    ELSIF ((x0 = FALSE) AND  (x1 = FALSE) AND  (x2 = TRUE) AND  (x3 = TRUE) AND  ( TRUE ) AND  ( TRUE )) OR ((x0 = FALSE) AND  (x1 = TRUE) AND  (x2 = FALSE) AND  (x3 = TRUE) AND  ( TRUE ) AND  ( TRUE )) OR ((x0 = FALSE) AND  (x1 = TRUE) AND  (x2 = TRUE) AND  ( TRUE ) AND  ( TRUE ) AND  ( TRUE )) OR ((x0 = TRUE) AND  ( TRUE ) AND  (x2 = FALSE) AND  (x3 = TRUE) AND  ( TRUE ) AND  ( TRUE )) OR ((x0 = TRUE) AND  ( TRUE ) AND  (x2 = TRUE) AND  ( TRUE ) AND  ( TRUE ) AND  ( TRUE )) THEN 
        cstate98 := 617; y0 := FALSE; y1 := FALSE; y2 := FALSE;  
    ELSIF ((x0 = FALSE) AND  (x1 = TRUE) AND  (x2 = FALSE) AND  (x3 = FALSE) AND  ( TRUE ) AND  (x5 = FALSE)) OR ((x0 = TRUE) AND  ( TRUE ) AND  (x2 = FALSE) AND  (x3 = FALSE) AND  ( TRUE ) AND  (x5 = FALSE)) THEN 
        cstate98 := 3204; y0 := TRUE; y1 := FALSE; y2 := FALSE;  
    ELSIF ((x0 = FALSE) AND  (x1 = TRUE) AND  (x2 = FALSE) AND  (x3 = FALSE) AND  ( TRUE ) AND  (x5 = TRUE)) OR ((x0 = TRUE) AND  ( TRUE ) AND  (x2 = FALSE) AND  (x3 = FALSE) AND  ( TRUE ) AND  (x5 = TRUE)) THEN 
        cstate98 := 1190; y0 := FALSE; y1 := FALSE; y2 := FALSE;  
    END_IF;
2212:
    IF ((x0 = FALSE) AND  (x1 = FALSE) AND  (x2 = FALSE) AND  (x3 = FALSE) AND  ( TRUE ) AND  (x5 = FALSE)) OR ((x0 = FALSE) AND  (x1 = FALSE) AND  (x2 = FALSE) AND  (x3 = TRUE) AND  (x4 = FALSE) AND  (x5 = FALSE)) THEN 
        cstate98 := 2212; y0 := FALSE; y1 := FALSE; y2 := FALSE;  
    ELSIF ((x0 = FALSE) AND  (x1 = FALSE) AND  (x2 = FALSE) AND  (x3 = FALSE) AND  ( TRUE ) AND  (x5 = TRUE)) OR ((x0 = FALSE) AND  (x1 = FALSE) AND  (x2 = FALSE) AND  (x3 = TRUE) AND  (x4 = FALSE) AND  (x5 = TRUE)) THEN 
        cstate98 := 2215; y0 := FALSE; y1 := FALSE; y2 := FALSE;  
    ELSIF ((x0 = FALSE) AND  (x1 = FALSE) AND  (x2 = FALSE) AND  (x3 = TRUE) AND  (x4 = TRUE) AND  (x5 = FALSE)) THEN 
        cstate98 := 236; y0 := FALSE; y1 := FALSE; y2 := TRUE;  
    ELSIF ((x0 = FALSE) AND  (x1 = FALSE) AND  (x2 = FALSE) AND  (x3 = TRUE) AND  (x4 = TRUE) AND  (x5 = TRUE)) THEN 
        cstate98 := 2190; y0 := FALSE; y1 := FALSE; y2 := FALSE;  
    ELSIF ((x0 = FALSE) AND  (x1 = FALSE) AND  (x2 = TRUE) AND  (x3 = FALSE) AND  ( TRUE ) AND  (x5 = FALSE)) THEN 
        cstate98 := 2704; y0 := FALSE; y1 := TRUE; y2 := FALSE;  
    ELSIF ((x0 = FALSE) AND  (x1 = FALSE) AND  (x2 = TRUE) AND  (x3 = FALSE) AND  ( TRUE ) AND  (x5 = TRUE)) THEN 
        cstate98 := 1714; y0 := FALSE; y1 := FALSE; y2 := FALSE;  
    ELSIF ((x0 = FALSE) AND  (x1 = FALSE) AND  (x2 = TRUE) AND  (x3 = TRUE) AND  ( TRUE ) AND  ( TRUE )) OR ((x0 = FALSE) AND  (x1 = TRUE) AND  (x2 = FALSE) AND  (x3 = TRUE) AND  ( TRUE ) AND  ( TRUE )) OR ((x0 = FALSE) AND  (x1 = TRUE) AND  (x2 = TRUE) AND  ( TRUE ) AND  ( TRUE ) AND  ( TRUE )) OR ((x0 = TRUE) AND  ( TRUE ) AND  (x2 = FALSE) AND  (x3 = TRUE) AND  ( TRUE ) AND  ( TRUE )) OR ((x0 = TRUE) AND  ( TRUE ) AND  (x2 = TRUE) AND  ( TRUE ) AND  ( TRUE ) AND  ( TRUE )) THEN 
        cstate98 := 617; y0 := FALSE; y1 := FALSE; y2 := FALSE;  
    ELSIF ((x0 = FALSE) AND  (x1 = TRUE) AND  (x2 = FALSE) AND  (x3 = FALSE) AND  ( TRUE ) AND  (x5 = FALSE)) OR ((x0 = TRUE) AND  ( TRUE ) AND  (x2 = FALSE) AND  (x3 = FALSE) AND  ( TRUE ) AND  (x5 = FALSE)) THEN 
        cstate98 := 3204; y0 := TRUE; y1 := FALSE; y2 := FALSE;  
    ELSIF ((x0 = FALSE) AND  (x1 = TRUE) AND  (x2 = FALSE) AND  (x3 = FALSE) AND  ( TRUE ) AND  (x5 = TRUE)) OR ((x0 = TRUE) AND  ( TRUE ) AND  (x2 = FALSE) AND  (x3 = FALSE) AND  ( TRUE ) AND  (x5 = TRUE)) THEN 
        cstate98 := 1190; y0 := FALSE; y1 := FALSE; y2 := FALSE;  
    END_IF;
236:
    IF ((x0 = FALSE) AND  (x1 = FALSE) AND  (x2 = FALSE) AND  (x3 = FALSE) AND  ( TRUE ) AND  (x5 = FALSE)) OR ((x0 = FALSE) AND  (x1 = FALSE) AND  (x2 = FALSE) AND  (x3 = TRUE) AND  (x4 = FALSE) AND  (x5 = FALSE)) OR ((x0 = FALSE) AND  (x1 = TRUE) AND  (x2 = FALSE) AND  (x3 = FALSE) AND  ( TRUE ) AND  (x5 = FALSE)) OR ((x0 = TRUE) AND  ( TRUE ) AND  (x2 = FALSE) AND  (x3 = FALSE) AND  ( TRUE ) AND  (x5 = FALSE)) THEN 
        cstate98 := 300; y0 := FALSE; y1 := FALSE; y2 := TRUE;  
    ELSIF ((x0 = FALSE) AND  (x1 = FALSE) AND  (x2 = FALSE) AND  (x3 = FALSE) AND  ( TRUE ) AND  (x5 = TRUE)) OR ((x0 = FALSE) AND  (x1 = FALSE) AND  (x2 = FALSE) AND  (x3 = TRUE) AND  (x4 = FALSE) AND  (x5 = TRUE)) THEN 
        cstate98 := 2223; y0 := FALSE; y1 := FALSE; y2 := FALSE;  
    ELSIF ((x0 = FALSE) AND  (x1 = FALSE) AND  (x2 = FALSE) AND  (x3 = TRUE) AND  (x4 = TRUE) AND  (x5 = FALSE)) THEN 
        cstate98 := 236; y0 := FALSE; y1 := FALSE; y2 := TRUE;  
    ELSIF ((x0 = FALSE) AND  (x1 = FALSE) AND  (x2 = FALSE) AND  (x3 = TRUE) AND  (x4 = TRUE) AND  (x5 = TRUE)) THEN 
        cstate98 := 2190; y0 := FALSE; y1 := FALSE; y2 := FALSE;  
    ELSIF ((x0 = FALSE) AND  (x1 = FALSE) AND  (x2 = TRUE) AND  (x3 = FALSE) AND  ( TRUE ) AND  (x5 = FALSE)) THEN 
        cstate98 := 296; y0 := FALSE; y1 := FALSE; y2 := TRUE;  
    ELSIF ((x0 = FALSE) AND  (x1 = FALSE) AND  (x2 = TRUE) AND  (x3 = FALSE) AND  ( TRUE ) AND  (x5 = TRUE)) THEN 
        cstate98 := 1706; y0 := FALSE; y1 := FALSE; y2 := FALSE;  
    ELSIF ((x0 = FALSE) AND  (x1 = FALSE) AND  (x2 = TRUE) AND  (x3 = TRUE) AND  ( TRUE ) AND  ( TRUE )) OR ((x0 = FALSE) AND  (x1 = TRUE) AND  (x2 = FALSE) AND  (x3 = TRUE) AND  ( TRUE ) AND  ( TRUE )) OR ((x0 = FALSE) AND  (x1 = TRUE) AND  (x2 = TRUE) AND  ( TRUE ) AND  ( TRUE ) AND  ( TRUE )) OR ((x0 = TRUE) AND  ( TRUE ) AND  (x2 = FALSE) AND  (x3 = TRUE) AND  ( TRUE ) AND  ( TRUE )) OR ((x0 = TRUE) AND  ( TRUE ) AND  (x2 = TRUE) AND  ( TRUE ) AND  ( TRUE ) AND  ( TRUE )) THEN 
        cstate98 := 617; y0 := FALSE; y1 := FALSE; y2 := FALSE;  
    ELSIF ((x0 = FALSE) AND  (x1 = TRUE) AND  (x2 = FALSE) AND  (x3 = FALSE) AND  ( TRUE ) AND  (x5 = TRUE)) OR ((x0 = TRUE) AND  ( TRUE ) AND  (x2 = FALSE) AND  (x3 = FALSE) AND  ( TRUE ) AND  (x5 = TRUE)) THEN 
        cstate98 := 1198; y0 := FALSE; y1 := FALSE; y2 := FALSE;  
    END_IF;
2214:
    IF ((x0 = FALSE) AND  (x1 = FALSE) AND  (x2 = FALSE) AND  (x3 = FALSE) AND  ( TRUE ) AND  (x5 = FALSE)) OR ((x0 = FALSE) AND  (x1 = FALSE) AND  (x2 = FALSE) AND  (x3 = TRUE) AND  (x4 = FALSE) AND  (x5 = FALSE)) THEN 
        cstate98 := 2214; y0 := FALSE; y1 := FALSE; y2 := FALSE;  
    ELSIF ((x0 = FALSE) AND  (x1 = FALSE) AND  (x2 = FALSE) AND  (x3 = FALSE) AND  ( TRUE ) AND  (x5 = TRUE)) OR ((x0 = FALSE) AND  (x1 = FALSE) AND  (x2 = FALSE) AND  (x3 = TRUE) AND  (x4 = FALSE) AND  (x5 = TRUE)) THEN 
        cstate98 := 2215; y0 := FALSE; y1 := FALSE; y2 := FALSE;  
    ELSIF ((x0 = FALSE) AND  (x1 = FALSE) AND  (x2 = FALSE) AND  (x3 = TRUE) AND  (x4 = TRUE) AND  (x5 = FALSE)) THEN 
        cstate98 := 238; y0 := FALSE; y1 := FALSE; y2 := TRUE;  
    ELSIF ((x0 = FALSE) AND  (x1 = FALSE) AND  (x2 = FALSE) AND  (x3 = TRUE) AND  (x4 = TRUE) AND  (x5 = TRUE)) THEN 
        cstate98 := 2190; y0 := FALSE; y1 := FALSE; y2 := FALSE;  
    ELSIF ((x0 = FALSE) AND  (x1 = FALSE) AND  (x2 = TRUE) AND  (x3 = FALSE) AND  ( TRUE ) AND  (x5 = FALSE)) THEN 
        cstate98 := 2706; y0 := FALSE; y1 := TRUE; y2 := FALSE;  
    ELSIF ((x0 = FALSE) AND  (x1 = FALSE) AND  (x2 = TRUE) AND  (x3 = FALSE) AND  ( TRUE ) AND  (x5 = TRUE)) THEN 
        cstate98 := 1714; y0 := FALSE; y1 := FALSE; y2 := FALSE;  
    ELSIF ((x0 = FALSE) AND  (x1 = FALSE) AND  (x2 = TRUE) AND  (x3 = TRUE) AND  ( TRUE ) AND  ( TRUE )) OR ((x0 = FALSE) AND  (x1 = TRUE) AND  (x2 = FALSE) AND  (x3 = TRUE) AND  ( TRUE ) AND  ( TRUE )) OR ((x0 = FALSE) AND  (x1 = TRUE) AND  (x2 = TRUE) AND  ( TRUE ) AND  ( TRUE ) AND  ( TRUE )) OR ((x0 = TRUE) AND  ( TRUE ) AND  (x2 = FALSE) AND  (x3 = TRUE) AND  ( TRUE ) AND  ( TRUE )) OR ((x0 = TRUE) AND  ( TRUE ) AND  (x2 = TRUE) AND  ( TRUE ) AND  ( TRUE ) AND  ( TRUE )) THEN 
        cstate98 := 617; y0 := FALSE; y1 := FALSE; y2 := FALSE;  
    ELSIF ((x0 = FALSE) AND  (x1 = TRUE) AND  (x2 = FALSE) AND  (x3 = FALSE) AND  ( TRUE ) AND  (x5 = FALSE)) OR ((x0 = TRUE) AND  ( TRUE ) AND  (x2 = FALSE) AND  (x3 = FALSE) AND  ( TRUE ) AND  (x5 = FALSE)) THEN 
        cstate98 := 3206; y0 := TRUE; y1 := FALSE; y2 := FALSE;  
    ELSIF ((x0 = FALSE) AND  (x1 = TRUE) AND  (x2 = FALSE) AND  (x3 = FALSE) AND  ( TRUE ) AND  (x5 = TRUE)) OR ((x0 = TRUE) AND  ( TRUE ) AND  (x2 = FALSE) AND  (x3 = FALSE) AND  ( TRUE ) AND  (x5 = TRUE)) THEN 
        cstate98 := 1190; y0 := FALSE; y1 := FALSE; y2 := FALSE;  
    END_IF;
238:
    IF ((x0 = FALSE) AND  (x1 = FALSE) AND  (x2 = FALSE) AND  (x3 = FALSE) AND  ( TRUE ) AND  (x5 = FALSE)) OR ((x0 = FALSE) AND  (x1 = FALSE) AND  (x2 = FALSE) AND  (x3 = TRUE) AND  (x4 = FALSE) AND  (x5 = FALSE)) OR ((x0 = FALSE) AND  (x1 = TRUE) AND  (x2 = FALSE) AND  (x3 = FALSE) AND  ( TRUE ) AND  (x5 = FALSE)) OR ((x0 = TRUE) AND  ( TRUE ) AND  (x2 = FALSE) AND  (x3 = FALSE) AND  ( TRUE ) AND  (x5 = FALSE)) THEN 
        cstate98 := 302; y0 := FALSE; y1 := FALSE; y2 := TRUE;  
    ELSIF ((x0 = FALSE) AND  (x1 = FALSE) AND  (x2 = FALSE) AND  (x3 = FALSE) AND  ( TRUE ) AND  (x5 = TRUE)) OR ((x0 = FALSE) AND  (x1 = FALSE) AND  (x2 = FALSE) AND  (x3 = TRUE) AND  (x4 = FALSE) AND  (x5 = TRUE)) THEN 
        cstate98 := 2223; y0 := FALSE; y1 := FALSE; y2 := FALSE;  
    ELSIF ((x0 = FALSE) AND  (x1 = FALSE) AND  (x2 = FALSE) AND  (x3 = TRUE) AND  (x4 = TRUE) AND  (x5 = FALSE)) THEN 
        cstate98 := 238; y0 := FALSE; y1 := FALSE; y2 := TRUE;  
    ELSIF ((x0 = FALSE) AND  (x1 = FALSE) AND  (x2 = FALSE) AND  (x3 = TRUE) AND  (x4 = TRUE) AND  (x5 = TRUE)) THEN 
        cstate98 := 2190; y0 := FALSE; y1 := FALSE; y2 := FALSE;  
    ELSIF ((x0 = FALSE) AND  (x1 = FALSE) AND  (x2 = TRUE) AND  (x3 = FALSE) AND  ( TRUE ) AND  (x5 = FALSE)) THEN 
        cstate98 := 298; y0 := FALSE; y1 := FALSE; y2 := TRUE;  
    ELSIF ((x0 = FALSE) AND  (x1 = FALSE) AND  (x2 = TRUE) AND  (x3 = FALSE) AND  ( TRUE ) AND  (x5 = TRUE)) THEN 
        cstate98 := 1706; y0 := FALSE; y1 := FALSE; y2 := FALSE;  
    ELSIF ((x0 = FALSE) AND  (x1 = FALSE) AND  (x2 = TRUE) AND  (x3 = TRUE) AND  ( TRUE ) AND  ( TRUE )) OR ((x0 = FALSE) AND  (x1 = TRUE) AND  (x2 = FALSE) AND  (x3 = TRUE) AND  ( TRUE ) AND  ( TRUE )) OR ((x0 = FALSE) AND  (x1 = TRUE) AND  (x2 = TRUE) AND  ( TRUE ) AND  ( TRUE ) AND  ( TRUE )) OR ((x0 = TRUE) AND  ( TRUE ) AND  (x2 = FALSE) AND  (x3 = TRUE) AND  ( TRUE ) AND  ( TRUE )) OR ((x0 = TRUE) AND  ( TRUE ) AND  (x2 = TRUE) AND  ( TRUE ) AND  ( TRUE ) AND  ( TRUE )) THEN 
        cstate98 := 617; y0 := FALSE; y1 := FALSE; y2 := FALSE;  
    ELSIF ((x0 = FALSE) AND  (x1 = TRUE) AND  (x2 = FALSE) AND  (x3 = FALSE) AND  ( TRUE ) AND  (x5 = TRUE)) OR ((x0 = TRUE) AND  ( TRUE ) AND  (x2 = FALSE) AND  (x3 = FALSE) AND  ( TRUE ) AND  (x5 = TRUE)) THEN 
        cstate98 := 1198; y0 := FALSE; y1 := FALSE; y2 := FALSE;  
    END_IF;
3210:
    IF ((x0 = FALSE) AND  (x1 = FALSE) AND  (x2 = FALSE) AND  ( TRUE ) AND  ( TRUE ) AND  (x5 = FALSE)) OR ((x0 = FALSE) AND  (x1 = FALSE) AND  (x2 = TRUE) AND  (x3 = FALSE) AND  ( TRUE ) AND  (x5 = FALSE)) THEN 
        cstate98 := 4234; y0 := TRUE; y1 := FALSE; y2 := FALSE;  
    ELSIF ((x0 = FALSE) AND  (x1 = FALSE) AND  (x2 = FALSE) AND  (x3 = FALSE) AND  ( TRUE ) AND  (x5 = TRUE)) OR ((x0 = FALSE) AND  (x1 = FALSE) AND  (x2 = FALSE) AND  (x3 = TRUE) AND  (x4 = FALSE) AND  (x5 = TRUE)) THEN 
        cstate98 := 2219; y0 := FALSE; y1 := FALSE; y2 := FALSE;  
    ELSIF ((x0 = FALSE) AND  (x1 = FALSE) AND  (x2 = FALSE) AND  (x3 = TRUE) AND  (x4 = TRUE) AND  (x5 = TRUE)) THEN 
        cstate98 := 2186; y0 := FALSE; y1 := FALSE; y2 := FALSE;  
    ELSIF ((x0 = FALSE) AND  (x1 = FALSE) AND  (x2 = TRUE) AND  (x3 = FALSE) AND  ( TRUE ) AND  (x5 = TRUE)) THEN 
        cstate98 := 1706; y0 := FALSE; y1 := FALSE; y2 := FALSE;  
    ELSIF ((x0 = FALSE) AND  (x1 = FALSE) AND  (x2 = TRUE) AND  (x3 = TRUE) AND  ( TRUE ) AND  ( TRUE )) OR ((x0 = FALSE) AND  (x1 = TRUE) AND  (x2 = FALSE) AND  (x3 = TRUE) AND  ( TRUE ) AND  ( TRUE )) OR ((x0 = FALSE) AND  (x1 = TRUE) AND  (x2 = TRUE) AND  ( TRUE ) AND  ( TRUE ) AND  ( TRUE )) OR ((x0 = TRUE) AND  ( TRUE ) AND  (x2 = FALSE) AND  (x3 = TRUE) AND  ( TRUE ) AND  ( TRUE )) OR ((x0 = TRUE) AND  ( TRUE ) AND  (x2 = TRUE) AND  ( TRUE ) AND  ( TRUE ) AND  ( TRUE )) THEN 
        cstate98 := 617; y0 := FALSE; y1 := FALSE; y2 := FALSE;  
    ELSIF ((x0 = FALSE) AND  (x1 = TRUE) AND  (x2 = FALSE) AND  (x3 = FALSE) AND  ( TRUE ) AND  (x5 = FALSE)) OR ((x0 = TRUE) AND  ( TRUE ) AND  (x2 = FALSE) AND  (x3 = FALSE) AND  ( TRUE ) AND  (x5 = FALSE)) THEN 
        cstate98 := 3210; y0 := TRUE; y1 := FALSE; y2 := FALSE;  
    ELSIF ((x0 = FALSE) AND  (x1 = TRUE) AND  (x2 = FALSE) AND  (x3 = FALSE) AND  ( TRUE ) AND  (x5 = TRUE)) OR ((x0 = TRUE) AND  ( TRUE ) AND  (x2 = FALSE) AND  (x3 = FALSE) AND  ( TRUE ) AND  (x5 = TRUE)) THEN 
        cstate98 := 1194; y0 := FALSE; y1 := FALSE; y2 := FALSE;  
    END_IF;
2119:
    IF ((x0 = FALSE) AND  (x1 = FALSE) AND  (x2 = FALSE) AND  (x3 = FALSE) AND  ( TRUE ) AND  ( TRUE )) OR ((x0 = FALSE) AND  (x1 = FALSE) AND  (x2 = FALSE) AND  (x3 = TRUE) AND  (x4 = FALSE) AND  ( TRUE )) THEN 
        cstate98 := 2119; y0 := FALSE; y1 := FALSE; y2 := FALSE;  
    ELSIF ((x0 = FALSE) AND  (x1 = FALSE) AND  (x2 = FALSE) AND  (x3 = TRUE) AND  (x4 = TRUE) AND  (x5 = FALSE)) THEN 
        cstate98 := 206; y0 := FALSE; y1 := FALSE; y2 := TRUE;  
    ELSIF ((x0 = FALSE) AND  (x1 = FALSE) AND  (x2 = FALSE) AND  (x3 = TRUE) AND  (x4 = TRUE) AND  (x5 = TRUE)) THEN 
        cstate98 := 2094; y0 := FALSE; y1 := FALSE; y2 := FALSE;  
    ELSIF ((x0 = FALSE) AND  (x1 = FALSE) AND  (x2 = TRUE) AND  (x3 = FALSE) AND  ( TRUE ) AND  (x5 = FALSE)) THEN 
        cstate98 := 2610; y0 := FALSE; y1 := TRUE; y2 := FALSE;  
    ELSIF ((x0 = FALSE) AND  (x1 = FALSE) AND  (x2 = TRUE) AND  (x3 = FALSE) AND  ( TRUE ) AND  (x5 = TRUE)) THEN 
        cstate98 := 1618; y0 := FALSE; y1 := FALSE; y2 := FALSE;  
    ELSIF ((x0 = FALSE) AND  (x1 = FALSE) AND  (x2 = TRUE) AND  (x3 = TRUE) AND  ( TRUE ) AND  ( TRUE )) OR ((x0 = FALSE) AND  (x1 = TRUE) AND  (x2 = FALSE) AND  (x3 = TRUE) AND  ( TRUE ) AND  ( TRUE )) OR ((x0 = FALSE) AND  (x1 = TRUE) AND  (x2 = TRUE) AND  ( TRUE ) AND  ( TRUE ) AND  ( TRUE )) OR ((x0 = TRUE) AND  ( TRUE ) AND  (x2 = FALSE) AND  (x3 = TRUE) AND  ( TRUE ) AND  ( TRUE )) OR ((x0 = TRUE) AND  ( TRUE ) AND  (x2 = TRUE) AND  ( TRUE ) AND  ( TRUE ) AND  ( TRUE )) THEN 
        cstate98 := 617; y0 := FALSE; y1 := FALSE; y2 := FALSE;  
    ELSIF ((x0 = FALSE) AND  (x1 = TRUE) AND  (x2 = FALSE) AND  (x3 = FALSE) AND  ( TRUE ) AND  (x5 = FALSE)) OR ((x0 = TRUE) AND  ( TRUE ) AND  (x2 = FALSE) AND  (x3 = FALSE) AND  ( TRUE ) AND  (x5 = FALSE)) THEN 
        cstate98 := 3206; y0 := TRUE; y1 := FALSE; y2 := FALSE;  
    ELSIF ((x0 = FALSE) AND  (x1 = TRUE) AND  (x2 = FALSE) AND  (x3 = FALSE) AND  ( TRUE ) AND  (x5 = TRUE)) OR ((x0 = TRUE) AND  ( TRUE ) AND  (x2 = FALSE) AND  (x3 = FALSE) AND  ( TRUE ) AND  (x5 = TRUE)) THEN 
        cstate98 := 1190; y0 := FALSE; y1 := FALSE; y2 := FALSE;  
    END_IF;
1610:
    IF ((x0 = FALSE) AND  (x1 = FALSE) AND  (x2 = FALSE) AND  (x3 = FALSE) AND  ( TRUE ) AND  (x5 = FALSE)) OR ((x0 = FALSE) AND  (x1 = FALSE) AND  (x2 = FALSE) AND  (x3 = TRUE) AND  (x4 = FALSE) AND  (x5 = FALSE)) THEN 
        cstate98 := 2122; y0 := FALSE; y1 := FALSE; y2 := FALSE;  
    ELSIF ((x0 = FALSE) AND  (x1 = FALSE) AND  (x2 = FALSE) AND  (x3 = FALSE) AND  ( TRUE ) AND  (x5 = TRUE)) OR ((x0 = FALSE) AND  (x1 = FALSE) AND  (x2 = FALSE) AND  (x3 = TRUE) AND  (x4 = FALSE) AND  (x5 = TRUE)) THEN 
        cstate98 := 2123; y0 := FALSE; y1 := FALSE; y2 := FALSE;  
    ELSIF ((x0 = FALSE) AND  (x1 = FALSE) AND  (x2 = FALSE) AND  (x3 = TRUE) AND  (x4 = TRUE) AND  (x5 = FALSE)) THEN 
        cstate98 := 202; y0 := FALSE; y1 := FALSE; y2 := TRUE;  
    ELSIF ((x0 = FALSE) AND  (x1 = FALSE) AND  (x2 = FALSE) AND  (x3 = TRUE) AND  (x4 = TRUE) AND  (x5 = TRUE)) THEN 
        cstate98 := 2090; y0 := FALSE; y1 := FALSE; y2 := FALSE;  
    ELSIF ((x0 = FALSE) AND  (x1 = FALSE) AND  (x2 = TRUE) AND  (x3 = FALSE) AND  ( TRUE ) AND  ( TRUE )) THEN 
        cstate98 := 1610; y0 := FALSE; y1 := FALSE; y2 := FALSE;  
    ELSIF ((x0 = FALSE) AND  (x1 = FALSE) AND  (x2 = TRUE) AND  (x3 = TRUE) AND  ( TRUE ) AND  ( TRUE )) OR ((x0 = FALSE) AND  (x1 = TRUE) AND  (x2 = FALSE) AND  (x3 = TRUE) AND  ( TRUE ) AND  ( TRUE )) OR ((x0 = FALSE) AND  (x1 = TRUE) AND  (x2 = TRUE) AND  ( TRUE ) AND  ( TRUE ) AND  ( TRUE )) OR ((x0 = TRUE) AND  ( TRUE ) AND  (x2 = FALSE) AND  (x3 = TRUE) AND  ( TRUE ) AND  ( TRUE )) OR ((x0 = TRUE) AND  ( TRUE ) AND  (x2 = TRUE) AND  ( TRUE ) AND  ( TRUE ) AND  ( TRUE )) THEN 
        cstate98 := 617; y0 := FALSE; y1 := FALSE; y2 := FALSE;  
    ELSIF ((x0 = FALSE) AND  (x1 = TRUE) AND  (x2 = FALSE) AND  (x3 = FALSE) AND  ( TRUE ) AND  (x5 = FALSE)) OR ((x0 = TRUE) AND  ( TRUE ) AND  (x2 = FALSE) AND  (x3 = FALSE) AND  ( TRUE ) AND  (x5 = FALSE)) THEN 
        cstate98 := 3210; y0 := TRUE; y1 := FALSE; y2 := FALSE;  
    ELSIF ((x0 = FALSE) AND  (x1 = TRUE) AND  (x2 = FALSE) AND  (x3 = FALSE) AND  ( TRUE ) AND  (x5 = TRUE)) OR ((x0 = TRUE) AND  ( TRUE ) AND  (x2 = FALSE) AND  (x3 = FALSE) AND  ( TRUE ) AND  (x5 = TRUE)) THEN 
        cstate98 := 1194; y0 := FALSE; y1 := FALSE; y2 := FALSE;  
    END_IF;
3218:
    IF ((x0 = FALSE) AND  (x1 = FALSE) AND  (x2 = FALSE) AND  (x3 = FALSE) AND  ( TRUE ) AND  (x5 = FALSE)) OR ((x0 = FALSE) AND  (x1 = FALSE) AND  (x2 = FALSE) AND  (x3 = TRUE) AND  (x4 = FALSE) AND  (x5 = FALSE)) OR ((x0 = FALSE) AND  (x1 = FALSE) AND  (x2 = TRUE) AND  (x3 = FALSE) AND  ( TRUE ) AND  (x5 = FALSE)) THEN 
        cstate98 := 4242; y0 := TRUE; y1 := FALSE; y2 := FALSE;  
    ELSIF ((x0 = FALSE) AND  (x1 = FALSE) AND  (x2 = FALSE) AND  (x3 = FALSE) AND  ( TRUE ) AND  (x5 = TRUE)) OR ((x0 = FALSE) AND  (x1 = FALSE) AND  (x2 = FALSE) AND  (x3 = TRUE) AND  (x4 = FALSE) AND  (x5 = TRUE)) THEN 
        cstate98 := 2227; y0 := FALSE; y1 := FALSE; y2 := FALSE;  
    ELSIF ((x0 = FALSE) AND  (x1 = FALSE) AND  (x2 = FALSE) AND  (x3 = TRUE) AND  (x4 = TRUE) AND  (x5 = FALSE)) THEN 
        cstate98 := 4234; y0 := TRUE; y1 := FALSE; y2 := FALSE;  
    ELSIF ((x0 = FALSE) AND  (x1 = FALSE) AND  (x2 = FALSE) AND  (x3 = TRUE) AND  (x4 = TRUE) AND  (x5 = TRUE)) THEN 
        cstate98 := 2186; y0 := FALSE; y1 := FALSE; y2 := FALSE;  
    ELSIF ((x0 = FALSE) AND  (x1 = FALSE) AND  (x2 = TRUE) AND  (x3 = FALSE) AND  ( TRUE ) AND  (x5 = TRUE)) THEN 
        cstate98 := 1714; y0 := FALSE; y1 := FALSE; y2 := FALSE;  
    ELSIF ((x0 = FALSE) AND  (x1 = FALSE) AND  (x2 = TRUE) AND  (x3 = TRUE) AND  ( TRUE ) AND  ( TRUE )) OR ((x0 = FALSE) AND  (x1 = TRUE) AND  (x2 = FALSE) AND  (x3 = TRUE) AND  ( TRUE ) AND  ( TRUE )) OR ((x0 = FALSE) AND  (x1 = TRUE) AND  (x2 = TRUE) AND  ( TRUE ) AND  ( TRUE ) AND  ( TRUE )) OR ((x0 = TRUE) AND  ( TRUE ) AND  (x2 = FALSE) AND  (x3 = TRUE) AND  ( TRUE ) AND  ( TRUE )) OR ((x0 = TRUE) AND  ( TRUE ) AND  (x2 = TRUE) AND  ( TRUE ) AND  ( TRUE ) AND  ( TRUE )) THEN 
        cstate98 := 617; y0 := FALSE; y1 := FALSE; y2 := FALSE;  
    ELSIF ((x0 = FALSE) AND  (x1 = TRUE) AND  (x2 = FALSE) AND  (x3 = FALSE) AND  ( TRUE ) AND  (x5 = FALSE)) OR ((x0 = TRUE) AND  ( TRUE ) AND  (x2 = FALSE) AND  (x3 = FALSE) AND  ( TRUE ) AND  (x5 = FALSE)) THEN 
        cstate98 := 3218; y0 := TRUE; y1 := FALSE; y2 := FALSE;  
    ELSIF ((x0 = FALSE) AND  (x1 = TRUE) AND  (x2 = FALSE) AND  (x3 = FALSE) AND  ( TRUE ) AND  (x5 = TRUE)) OR ((x0 = TRUE) AND  ( TRUE ) AND  (x2 = FALSE) AND  (x3 = FALSE) AND  ( TRUE ) AND  (x5 = TRUE)) THEN 
        cstate98 := 1202; y0 := FALSE; y1 := FALSE; y2 := FALSE;  
    END_IF;
3216:
    IF ((x0 = FALSE) AND  (x1 = FALSE) AND  (x2 = FALSE) AND  (x3 = FALSE) AND  ( TRUE ) AND  (x5 = FALSE)) OR ((x0 = FALSE) AND  (x1 = FALSE) AND  (x2 = FALSE) AND  (x3 = TRUE) AND  (x4 = FALSE) AND  (x5 = FALSE)) OR ((x0 = FALSE) AND  (x1 = FALSE) AND  (x2 = TRUE) AND  (x3 = FALSE) AND  ( TRUE ) AND  (x5 = FALSE)) THEN 
        cstate98 := 4240; y0 := TRUE; y1 := FALSE; y2 := FALSE;  
    ELSIF ((x0 = FALSE) AND  (x1 = FALSE) AND  (x2 = FALSE) AND  (x3 = FALSE) AND  ( TRUE ) AND  (x5 = TRUE)) OR ((x0 = FALSE) AND  (x1 = FALSE) AND  (x2 = FALSE) AND  (x3 = TRUE) AND  (x4 = FALSE) AND  (x5 = TRUE)) THEN 
        cstate98 := 2227; y0 := FALSE; y1 := FALSE; y2 := FALSE;  
    ELSIF ((x0 = FALSE) AND  (x1 = FALSE) AND  (x2 = FALSE) AND  (x3 = TRUE) AND  (x4 = TRUE) AND  (x5 = FALSE)) THEN 
        cstate98 := 4232; y0 := TRUE; y1 := FALSE; y2 := FALSE;  
    ELSIF ((x0 = FALSE) AND  (x1 = FALSE) AND  (x2 = FALSE) AND  (x3 = TRUE) AND  (x4 = TRUE) AND  (x5 = TRUE)) THEN 
        cstate98 := 2186; y0 := FALSE; y1 := FALSE; y2 := FALSE;  
    ELSIF ((x0 = FALSE) AND  (x1 = FALSE) AND  (x2 = TRUE) AND  (x3 = FALSE) AND  ( TRUE ) AND  (x5 = TRUE)) THEN 
        cstate98 := 1714; y0 := FALSE; y1 := FALSE; y2 := FALSE;  
    ELSIF ((x0 = FALSE) AND  (x1 = FALSE) AND  (x2 = TRUE) AND  (x3 = TRUE) AND  ( TRUE ) AND  ( TRUE )) OR ((x0 = FALSE) AND  (x1 = TRUE) AND  (x2 = FALSE) AND  (x3 = TRUE) AND  ( TRUE ) AND  ( TRUE )) OR ((x0 = FALSE) AND  (x1 = TRUE) AND  (x2 = TRUE) AND  ( TRUE ) AND  ( TRUE ) AND  ( TRUE )) OR ((x0 = TRUE) AND  ( TRUE ) AND  (x2 = FALSE) AND  (x3 = TRUE) AND  ( TRUE ) AND  ( TRUE )) OR ((x0 = TRUE) AND  ( TRUE ) AND  (x2 = TRUE) AND  ( TRUE ) AND  ( TRUE ) AND  ( TRUE )) THEN 
        cstate98 := 617; y0 := FALSE; y1 := FALSE; y2 := FALSE;  
    ELSIF ((x0 = FALSE) AND  (x1 = TRUE) AND  (x2 = FALSE) AND  (x3 = FALSE) AND  ( TRUE ) AND  (x5 = FALSE)) OR ((x0 = TRUE) AND  ( TRUE ) AND  (x2 = FALSE) AND  (x3 = FALSE) AND  ( TRUE ) AND  (x5 = FALSE)) THEN 
        cstate98 := 3216; y0 := TRUE; y1 := FALSE; y2 := FALSE;  
    ELSIF ((x0 = FALSE) AND  (x1 = TRUE) AND  (x2 = FALSE) AND  (x3 = FALSE) AND  ( TRUE ) AND  (x5 = TRUE)) OR ((x0 = TRUE) AND  ( TRUE ) AND  (x2 = FALSE) AND  (x3 = FALSE) AND  ( TRUE ) AND  (x5 = TRUE)) THEN 
        cstate98 := 1202; y0 := FALSE; y1 := FALSE; y2 := FALSE;  
    END_IF;
2131:
    IF ((x0 = FALSE) AND  (x1 = FALSE) AND  (x2 = FALSE) AND  (x3 = FALSE) AND  ( TRUE ) AND  ( TRUE )) OR ((x0 = FALSE) AND  (x1 = FALSE) AND  (x2 = FALSE) AND  (x3 = TRUE) AND  (x4 = FALSE) AND  ( TRUE )) THEN 
        cstate98 := 2131; y0 := FALSE; y1 := FALSE; y2 := FALSE;  
    ELSIF ((x0 = FALSE) AND  (x1 = FALSE) AND  (x2 = FALSE) AND  (x3 = TRUE) AND  (x4 = TRUE) AND  (x5 = FALSE)) THEN 
        cstate98 := 202; y0 := FALSE; y1 := FALSE; y2 := TRUE;  
    ELSIF ((x0 = FALSE) AND  (x1 = FALSE) AND  (x2 = FALSE) AND  (x3 = TRUE) AND  (x4 = TRUE) AND  (x5 = TRUE)) THEN 
        cstate98 := 2090; y0 := FALSE; y1 := FALSE; y2 := FALSE;  
    ELSIF ((x0 = FALSE) AND  (x1 = FALSE) AND  (x2 = TRUE) AND  (x3 = FALSE) AND  ( TRUE ) AND  (x5 = FALSE)) THEN 
        cstate98 := 2610; y0 := FALSE; y1 := TRUE; y2 := FALSE;  
    ELSIF ((x0 = FALSE) AND  (x1 = FALSE) AND  (x2 = TRUE) AND  (x3 = FALSE) AND  ( TRUE ) AND  (x5 = TRUE)) THEN 
        cstate98 := 1618; y0 := FALSE; y1 := FALSE; y2 := FALSE;  
    ELSIF ((x0 = FALSE) AND  (x1 = FALSE) AND  (x2 = TRUE) AND  (x3 = TRUE) AND  ( TRUE ) AND  ( TRUE )) OR ((x0 = FALSE) AND  (x1 = TRUE) AND  (x2 = FALSE) AND  (x3 = TRUE) AND  ( TRUE ) AND  ( TRUE )) OR ((x0 = FALSE) AND  (x1 = TRUE) AND  (x2 = TRUE) AND  ( TRUE ) AND  ( TRUE ) AND  ( TRUE )) OR ((x0 = TRUE) AND  ( TRUE ) AND  (x2 = FALSE) AND  (x3 = TRUE) AND  ( TRUE ) AND  ( TRUE )) OR ((x0 = TRUE) AND  ( TRUE ) AND  (x2 = TRUE) AND  ( TRUE ) AND  ( TRUE ) AND  ( TRUE )) THEN 
        cstate98 := 617; y0 := FALSE; y1 := FALSE; y2 := FALSE;  
    ELSIF ((x0 = FALSE) AND  (x1 = TRUE) AND  (x2 = FALSE) AND  (x3 = FALSE) AND  ( TRUE ) AND  (x5 = FALSE)) OR ((x0 = TRUE) AND  ( TRUE ) AND  (x2 = FALSE) AND  (x3 = FALSE) AND  ( TRUE ) AND  (x5 = FALSE)) THEN 
        cstate98 := 3218; y0 := TRUE; y1 := FALSE; y2 := FALSE;  
    ELSIF ((x0 = FALSE) AND  (x1 = TRUE) AND  (x2 = FALSE) AND  (x3 = FALSE) AND  ( TRUE ) AND  (x5 = TRUE)) OR ((x0 = TRUE) AND  ( TRUE ) AND  (x2 = FALSE) AND  (x3 = FALSE) AND  ( TRUE ) AND  (x5 = TRUE)) THEN 
        cstate98 := 1202; y0 := FALSE; y1 := FALSE; y2 := FALSE;  
    END_IF;
2130:
    IF ((x0 = FALSE) AND  (x1 = FALSE) AND  (x2 = FALSE) AND  (x3 = FALSE) AND  ( TRUE ) AND  (x5 = FALSE)) OR ((x0 = FALSE) AND  (x1 = FALSE) AND  (x2 = FALSE) AND  (x3 = TRUE) AND  (x4 = FALSE) AND  (x5 = FALSE)) THEN 
        cstate98 := 2130; y0 := FALSE; y1 := FALSE; y2 := FALSE;  
    ELSIF ((x0 = FALSE) AND  (x1 = FALSE) AND  (x2 = FALSE) AND  (x3 = FALSE) AND  ( TRUE ) AND  (x5 = TRUE)) OR ((x0 = FALSE) AND  (x1 = FALSE) AND  (x2 = FALSE) AND  (x3 = TRUE) AND  (x4 = FALSE) AND  (x5 = TRUE)) THEN 
        cstate98 := 2131; y0 := FALSE; y1 := FALSE; y2 := FALSE;  
    ELSIF ((x0 = FALSE) AND  (x1 = FALSE) AND  (x2 = FALSE) AND  (x3 = TRUE) AND  (x4 = TRUE) AND  (x5 = FALSE)) THEN 
        cstate98 := 202; y0 := FALSE; y1 := FALSE; y2 := TRUE;  
    ELSIF ((x0 = FALSE) AND  (x1 = FALSE) AND  (x2 = FALSE) AND  (x3 = TRUE) AND  (x4 = TRUE) AND  (x5 = TRUE)) THEN 
        cstate98 := 2090; y0 := FALSE; y1 := FALSE; y2 := FALSE;  
    ELSIF ((x0 = FALSE) AND  (x1 = FALSE) AND  (x2 = TRUE) AND  (x3 = FALSE) AND  ( TRUE ) AND  (x5 = FALSE)) THEN 
        cstate98 := 2610; y0 := FALSE; y1 := TRUE; y2 := FALSE;  
    ELSIF ((x0 = FALSE) AND  (x1 = FALSE) AND  (x2 = TRUE) AND  (x3 = FALSE) AND  ( TRUE ) AND  (x5 = TRUE)) THEN 
        cstate98 := 1618; y0 := FALSE; y1 := FALSE; y2 := FALSE;  
    ELSIF ((x0 = FALSE) AND  (x1 = FALSE) AND  (x2 = TRUE) AND  (x3 = TRUE) AND  ( TRUE ) AND  ( TRUE )) OR ((x0 = FALSE) AND  (x1 = TRUE) AND  (x2 = FALSE) AND  (x3 = TRUE) AND  ( TRUE ) AND  ( TRUE )) OR ((x0 = FALSE) AND  (x1 = TRUE) AND  (x2 = TRUE) AND  ( TRUE ) AND  ( TRUE ) AND  ( TRUE )) OR ((x0 = TRUE) AND  ( TRUE ) AND  (x2 = FALSE) AND  (x3 = TRUE) AND  ( TRUE ) AND  ( TRUE )) OR ((x0 = TRUE) AND  ( TRUE ) AND  (x2 = TRUE) AND  ( TRUE ) AND  ( TRUE ) AND  ( TRUE )) THEN 
        cstate98 := 617; y0 := FALSE; y1 := FALSE; y2 := FALSE;  
    ELSIF ((x0 = FALSE) AND  (x1 = TRUE) AND  (x2 = FALSE) AND  (x3 = FALSE) AND  ( TRUE ) AND  (x5 = FALSE)) OR ((x0 = TRUE) AND  ( TRUE ) AND  (x2 = FALSE) AND  (x3 = FALSE) AND  ( TRUE ) AND  (x5 = FALSE)) THEN 
        cstate98 := 3218; y0 := TRUE; y1 := FALSE; y2 := FALSE;  
    ELSIF ((x0 = FALSE) AND  (x1 = TRUE) AND  (x2 = FALSE) AND  (x3 = FALSE) AND  ( TRUE ) AND  (x5 = TRUE)) OR ((x0 = TRUE) AND  ( TRUE ) AND  (x2 = FALSE) AND  (x3 = FALSE) AND  ( TRUE ) AND  (x5 = TRUE)) THEN 
        cstate98 := 1202; y0 := FALSE; y1 := FALSE; y2 := FALSE;  
    END_IF;
3214:
    IF ((x0 = FALSE) AND  (x1 = FALSE) AND  (x2 = FALSE) AND  ( TRUE ) AND  ( TRUE ) AND  (x5 = FALSE)) THEN 
        cstate98 := 4238; y0 := TRUE; y1 := FALSE; y2 := FALSE;  
    ELSIF ((x0 = FALSE) AND  (x1 = FALSE) AND  (x2 = FALSE) AND  (x3 = FALSE) AND  ( TRUE ) AND  (x5 = TRUE)) OR ((x0 = FALSE) AND  (x1 = FALSE) AND  (x2 = FALSE) AND  (x3 = TRUE) AND  (x4 = FALSE) AND  (x5 = TRUE)) THEN 
        cstate98 := 2223; y0 := FALSE; y1 := FALSE; y2 := FALSE;  
    ELSIF ((x0 = FALSE) AND  (x1 = FALSE) AND  (x2 = FALSE) AND  (x3 = TRUE) AND  (x4 = TRUE) AND  (x5 = TRUE)) THEN 
        cstate98 := 2190; y0 := FALSE; y1 := FALSE; y2 := FALSE;  
    ELSIF ((x0 = FALSE) AND  (x1 = FALSE) AND  (x2 = TRUE) AND  (x3 = FALSE) AND  ( TRUE ) AND  (x5 = FALSE)) THEN 
        cstate98 := 4234; y0 := TRUE; y1 := FALSE; y2 := FALSE;  
    ELSIF ((x0 = FALSE) AND  (x1 = FALSE) AND  (x2 = TRUE) AND  (x3 = FALSE) AND  ( TRUE ) AND  (x5 = TRUE)) THEN 
        cstate98 := 1706; y0 := FALSE; y1 := FALSE; y2 := FALSE;  
    ELSIF ((x0 = FALSE) AND  (x1 = FALSE) AND  (x2 = TRUE) AND  (x3 = TRUE) AND  ( TRUE ) AND  ( TRUE )) OR ((x0 = FALSE) AND  (x1 = TRUE) AND  (x2 = FALSE) AND  (x3 = TRUE) AND  ( TRUE ) AND  ( TRUE )) OR ((x0 = FALSE) AND  (x1 = TRUE) AND  (x2 = TRUE) AND  ( TRUE ) AND  ( TRUE ) AND  ( TRUE )) OR ((x0 = TRUE) AND  ( TRUE ) AND  (x2 = FALSE) AND  (x3 = TRUE) AND  ( TRUE ) AND  ( TRUE )) OR ((x0 = TRUE) AND  ( TRUE ) AND  (x2 = TRUE) AND  ( TRUE ) AND  ( TRUE ) AND  ( TRUE )) THEN 
        cstate98 := 617; y0 := FALSE; y1 := FALSE; y2 := FALSE;  
    ELSIF ((x0 = FALSE) AND  (x1 = TRUE) AND  (x2 = FALSE) AND  (x3 = FALSE) AND  ( TRUE ) AND  (x5 = FALSE)) OR ((x0 = TRUE) AND  ( TRUE ) AND  (x2 = FALSE) AND  (x3 = FALSE) AND  ( TRUE ) AND  (x5 = FALSE)) THEN 
        cstate98 := 3214; y0 := TRUE; y1 := FALSE; y2 := FALSE;  
    ELSIF ((x0 = FALSE) AND  (x1 = TRUE) AND  (x2 = FALSE) AND  (x3 = FALSE) AND  ( TRUE ) AND  (x5 = TRUE)) OR ((x0 = TRUE) AND  ( TRUE ) AND  (x2 = FALSE) AND  (x3 = FALSE) AND  ( TRUE ) AND  (x5 = TRUE)) THEN 
        cstate98 := 1198; y0 := FALSE; y1 := FALSE; y2 := FALSE;  
    END_IF;
4228:
    IF ((x0 = FALSE) AND  (x1 = FALSE) AND  (x2 = FALSE) AND  (x3 = FALSE) AND  ( TRUE ) AND  (x5 = FALSE)) OR ((x0 = FALSE) AND  (x1 = FALSE) AND  (x2 = FALSE) AND  (x3 = TRUE) AND  (x4 = FALSE) AND  (x5 = FALSE)) THEN 
        cstate98 := 4228; y0 := TRUE; y1 := FALSE; y2 := FALSE;  
    ELSIF ((x0 = FALSE) AND  (x1 = FALSE) AND  (x2 = FALSE) AND  (x3 = FALSE) AND  ( TRUE ) AND  (x5 = TRUE)) OR ((x0 = FALSE) AND  (x1 = FALSE) AND  (x2 = FALSE) AND  (x3 = TRUE) AND  (x4 = FALSE) AND  (x5 = TRUE)) THEN 
        cstate98 := 2215; y0 := FALSE; y1 := FALSE; y2 := FALSE;  
    ELSIF ((x0 = FALSE) AND  (x1 = FALSE) AND  (x2 = FALSE) AND  (x3 = TRUE) AND  (x4 = TRUE) AND  (x5 = FALSE)) THEN 
        cstate98 := 4236; y0 := TRUE; y1 := FALSE; y2 := FALSE;  
    ELSIF ((x0 = FALSE) AND  (x1 = FALSE) AND  (x2 = FALSE) AND  (x3 = TRUE) AND  (x4 = TRUE) AND  (x5 = TRUE)) THEN 
        cstate98 := 2190; y0 := FALSE; y1 := FALSE; y2 := FALSE;  
    ELSIF ((x0 = FALSE) AND  (x1 = FALSE) AND  (x2 = TRUE) AND  (x3 = FALSE) AND  ( TRUE ) AND  (x5 = FALSE)) THEN 
        cstate98 := 4240; y0 := TRUE; y1 := FALSE; y2 := FALSE;  
    ELSIF ((x0 = FALSE) AND  (x1 = FALSE) AND  (x2 = TRUE) AND  (x3 = FALSE) AND  ( TRUE ) AND  (x5 = TRUE)) THEN 
        cstate98 := 1714; y0 := FALSE; y1 := FALSE; y2 := FALSE;  
    ELSIF ((x0 = FALSE) AND  (x1 = FALSE) AND  (x2 = TRUE) AND  (x3 = TRUE) AND  ( TRUE ) AND  ( TRUE )) OR ((x0 = FALSE) AND  (x1 = TRUE) AND  (x2 = FALSE) AND  (x3 = TRUE) AND  ( TRUE ) AND  ( TRUE )) OR ((x0 = FALSE) AND  (x1 = TRUE) AND  (x2 = TRUE) AND  ( TRUE ) AND  ( TRUE ) AND  ( TRUE )) OR ((x0 = TRUE) AND  ( TRUE ) AND  (x2 = FALSE) AND  (x3 = TRUE) AND  ( TRUE ) AND  ( TRUE )) OR ((x0 = TRUE) AND  ( TRUE ) AND  (x2 = TRUE) AND  ( TRUE ) AND  ( TRUE ) AND  ( TRUE )) THEN 
        cstate98 := 617; y0 := FALSE; y1 := FALSE; y2 := FALSE;  
    ELSIF ((x0 = FALSE) AND  (x1 = TRUE) AND  (x2 = FALSE) AND  (x3 = FALSE) AND  ( TRUE ) AND  (x5 = FALSE)) OR ((x0 = TRUE) AND  ( TRUE ) AND  (x2 = FALSE) AND  (x3 = FALSE) AND  ( TRUE ) AND  (x5 = FALSE)) THEN 
        cstate98 := 3204; y0 := TRUE; y1 := FALSE; y2 := FALSE;  
    ELSIF ((x0 = FALSE) AND  (x1 = TRUE) AND  (x2 = FALSE) AND  (x3 = FALSE) AND  ( TRUE ) AND  (x5 = TRUE)) OR ((x0 = TRUE) AND  ( TRUE ) AND  (x2 = FALSE) AND  (x3 = FALSE) AND  ( TRUE ) AND  (x5 = TRUE)) THEN 
        cstate98 := 1190; y0 := FALSE; y1 := FALSE; y2 := FALSE;  
    END_IF;
3212:
    IF ((x0 = FALSE) AND  (x1 = FALSE) AND  (x2 = FALSE) AND  ( TRUE ) AND  ( TRUE ) AND  (x5 = FALSE)) THEN 
        cstate98 := 4236; y0 := TRUE; y1 := FALSE; y2 := FALSE;  
    ELSIF ((x0 = FALSE) AND  (x1 = FALSE) AND  (x2 = FALSE) AND  (x3 = FALSE) AND  ( TRUE ) AND  (x5 = TRUE)) OR ((x0 = FALSE) AND  (x1 = FALSE) AND  (x2 = FALSE) AND  (x3 = TRUE) AND  (x4 = FALSE) AND  (x5 = TRUE)) THEN 
        cstate98 := 2223; y0 := FALSE; y1 := FALSE; y2 := FALSE;  
    ELSIF ((x0 = FALSE) AND  (x1 = FALSE) AND  (x2 = FALSE) AND  (x3 = TRUE) AND  (x4 = TRUE) AND  (x5 = TRUE)) THEN 
        cstate98 := 2190; y0 := FALSE; y1 := FALSE; y2 := FALSE;  
    ELSIF ((x0 = FALSE) AND  (x1 = FALSE) AND  (x2 = TRUE) AND  (x3 = FALSE) AND  ( TRUE ) AND  (x5 = FALSE)) THEN 
        cstate98 := 4232; y0 := TRUE; y1 := FALSE; y2 := FALSE;  
    ELSIF ((x0 = FALSE) AND  (x1 = FALSE) AND  (x2 = TRUE) AND  (x3 = FALSE) AND  ( TRUE ) AND  (x5 = TRUE)) THEN 
        cstate98 := 1706; y0 := FALSE; y1 := FALSE; y2 := FALSE;  
    ELSIF ((x0 = FALSE) AND  (x1 = FALSE) AND  (x2 = TRUE) AND  (x3 = TRUE) AND  ( TRUE ) AND  ( TRUE )) OR ((x0 = FALSE) AND  (x1 = TRUE) AND  (x2 = FALSE) AND  (x3 = TRUE) AND  ( TRUE ) AND  ( TRUE )) OR ((x0 = FALSE) AND  (x1 = TRUE) AND  (x2 = TRUE) AND  ( TRUE ) AND  ( TRUE ) AND  ( TRUE )) OR ((x0 = TRUE) AND  ( TRUE ) AND  (x2 = FALSE) AND  (x3 = TRUE) AND  ( TRUE ) AND  ( TRUE )) OR ((x0 = TRUE) AND  ( TRUE ) AND  (x2 = TRUE) AND  ( TRUE ) AND  ( TRUE ) AND  ( TRUE )) THEN 
        cstate98 := 617; y0 := FALSE; y1 := FALSE; y2 := FALSE;  
    ELSIF ((x0 = FALSE) AND  (x1 = TRUE) AND  (x2 = FALSE) AND  (x3 = FALSE) AND  ( TRUE ) AND  (x5 = FALSE)) OR ((x0 = TRUE) AND  ( TRUE ) AND  (x2 = FALSE) AND  (x3 = FALSE) AND  ( TRUE ) AND  (x5 = FALSE)) THEN 
        cstate98 := 3212; y0 := TRUE; y1 := FALSE; y2 := FALSE;  
    ELSIF ((x0 = FALSE) AND  (x1 = TRUE) AND  (x2 = FALSE) AND  (x3 = FALSE) AND  ( TRUE ) AND  (x5 = TRUE)) OR ((x0 = TRUE) AND  ( TRUE ) AND  (x2 = FALSE) AND  (x3 = FALSE) AND  ( TRUE ) AND  (x5 = TRUE)) THEN 
        cstate98 := 1198; y0 := FALSE; y1 := FALSE; y2 := FALSE;  
    END_IF;
2698:
    IF ((x0 = FALSE) AND  (x1 = FALSE) AND  (x2 = FALSE) AND  ( TRUE ) AND  ( TRUE ) AND  (x5 = FALSE)) OR ((x0 = FALSE) AND  (x1 = TRUE) AND  (x2 = FALSE) AND  (x3 = FALSE) AND  ( TRUE ) AND  (x5 = FALSE)) OR ((x0 = TRUE) AND  ( TRUE ) AND  (x2 = FALSE) AND  (x3 = FALSE) AND  ( TRUE ) AND  (x5 = FALSE)) THEN 
        cstate98 := 3722; y0 := FALSE; y1 := TRUE; y2 := FALSE;  
    ELSIF ((x0 = FALSE) AND  (x1 = FALSE) AND  (x2 = FALSE) AND  (x3 = FALSE) AND  ( TRUE ) AND  (x5 = TRUE)) OR ((x0 = FALSE) AND  (x1 = FALSE) AND  (x2 = FALSE) AND  (x3 = TRUE) AND  (x4 = FALSE) AND  (x5 = TRUE)) THEN 
        cstate98 := 2219; y0 := FALSE; y1 := FALSE; y2 := FALSE;  
    ELSIF ((x0 = FALSE) AND  (x1 = FALSE) AND  (x2 = FALSE) AND  (x3 = TRUE) AND  (x4 = TRUE) AND  (x5 = TRUE)) THEN 
        cstate98 := 2186; y0 := FALSE; y1 := FALSE; y2 := FALSE;  
    ELSIF ((x0 = FALSE) AND  (x1 = FALSE) AND  (x2 = TRUE) AND  (x3 = FALSE) AND  ( TRUE ) AND  (x5 = FALSE)) THEN 
        cstate98 := 2698; y0 := FALSE; y1 := TRUE; y2 := FALSE;  
    ELSIF ((x0 = FALSE) AND  (x1 = FALSE) AND  (x2 = TRUE) AND  (x3 = FALSE) AND  ( TRUE ) AND  (x5 = TRUE)) THEN 
        cstate98 := 1706; y0 := FALSE; y1 := FALSE; y2 := FALSE;  
    ELSIF ((x0 = FALSE) AND  (x1 = FALSE) AND  (x2 = TRUE) AND  (x3 = TRUE) AND  ( TRUE ) AND  ( TRUE )) OR ((x0 = FALSE) AND  (x1 = TRUE) AND  (x2 = FALSE) AND  (x3 = TRUE) AND  ( TRUE ) AND  ( TRUE )) OR ((x0 = FALSE) AND  (x1 = TRUE) AND  (x2 = TRUE) AND  ( TRUE ) AND  ( TRUE ) AND  ( TRUE )) OR ((x0 = TRUE) AND  ( TRUE ) AND  (x2 = FALSE) AND  (x3 = TRUE) AND  ( TRUE ) AND  ( TRUE )) OR ((x0 = TRUE) AND  ( TRUE ) AND  (x2 = TRUE) AND  ( TRUE ) AND  ( TRUE ) AND  ( TRUE )) THEN 
        cstate98 := 617; y0 := FALSE; y1 := FALSE; y2 := FALSE;  
    ELSIF ((x0 = FALSE) AND  (x1 = TRUE) AND  (x2 = FALSE) AND  (x3 = FALSE) AND  ( TRUE ) AND  (x5 = TRUE)) OR ((x0 = TRUE) AND  ( TRUE ) AND  (x2 = FALSE) AND  (x3 = FALSE) AND  ( TRUE ) AND  (x5 = TRUE)) THEN 
        cstate98 := 1194; y0 := FALSE; y1 := FALSE; y2 := FALSE;  
    END_IF;
2222:
    IF ((x0 = FALSE) AND  (x1 = FALSE) AND  (x2 = FALSE) AND  (x3 = FALSE) AND  ( TRUE ) AND  (x5 = FALSE)) OR ((x0 = FALSE) AND  (x1 = FALSE) AND  (x2 = FALSE) AND  (x3 = TRUE) AND  (x4 = FALSE) AND  (x5 = FALSE)) THEN 
        cstate98 := 2222; y0 := FALSE; y1 := FALSE; y2 := FALSE;  
    ELSIF ((x0 = FALSE) AND  (x1 = FALSE) AND  (x2 = FALSE) AND  (x3 = FALSE) AND  ( TRUE ) AND  (x5 = TRUE)) OR ((x0 = FALSE) AND  (x1 = FALSE) AND  (x2 = FALSE) AND  (x3 = TRUE) AND  (x4 = FALSE) AND  (x5 = TRUE)) THEN 
        cstate98 := 2223; y0 := FALSE; y1 := FALSE; y2 := FALSE;  
    ELSIF ((x0 = FALSE) AND  (x1 = FALSE) AND  (x2 = FALSE) AND  (x3 = TRUE) AND  (x4 = TRUE) AND  (x5 = FALSE)) THEN 
        cstate98 := 238; y0 := FALSE; y1 := FALSE; y2 := TRUE;  
    ELSIF ((x0 = FALSE) AND  (x1 = FALSE) AND  (x2 = FALSE) AND  (x3 = TRUE) AND  (x4 = TRUE) AND  (x5 = TRUE)) THEN 
        cstate98 := 2190; y0 := FALSE; y1 := FALSE; y2 := FALSE;  
    ELSIF ((x0 = FALSE) AND  (x1 = FALSE) AND  (x2 = TRUE) AND  (x3 = FALSE) AND  ( TRUE ) AND  (x5 = FALSE)) THEN 
        cstate98 := 2698; y0 := FALSE; y1 := TRUE; y2 := FALSE;  
    ELSIF ((x0 = FALSE) AND  (x1 = FALSE) AND  (x2 = TRUE) AND  (x3 = FALSE) AND  ( TRUE ) AND  (x5 = TRUE)) THEN 
        cstate98 := 1706; y0 := FALSE; y1 := FALSE; y2 := FALSE;  
    ELSIF ((x0 = FALSE) AND  (x1 = FALSE) AND  (x2 = TRUE) AND  (x3 = TRUE) AND  ( TRUE ) AND  ( TRUE )) OR ((x0 = FALSE) AND  (x1 = TRUE) AND  (x2 = FALSE) AND  (x3 = TRUE) AND  ( TRUE ) AND  ( TRUE )) OR ((x0 = FALSE) AND  (x1 = TRUE) AND  (x2 = TRUE) AND  ( TRUE ) AND  ( TRUE ) AND  ( TRUE )) OR ((x0 = TRUE) AND  ( TRUE ) AND  (x2 = FALSE) AND  (x3 = TRUE) AND  ( TRUE ) AND  ( TRUE )) OR ((x0 = TRUE) AND  ( TRUE ) AND  (x2 = TRUE) AND  ( TRUE ) AND  ( TRUE ) AND  ( TRUE )) THEN 
        cstate98 := 617; y0 := FALSE; y1 := FALSE; y2 := FALSE;  
    ELSIF ((x0 = FALSE) AND  (x1 = TRUE) AND  (x2 = FALSE) AND  (x3 = FALSE) AND  ( TRUE ) AND  (x5 = FALSE)) OR ((x0 = TRUE) AND  ( TRUE ) AND  (x2 = FALSE) AND  (x3 = FALSE) AND  ( TRUE ) AND  (x5 = FALSE)) THEN 
        cstate98 := 3214; y0 := TRUE; y1 := FALSE; y2 := FALSE;  
    ELSIF ((x0 = FALSE) AND  (x1 = TRUE) AND  (x2 = FALSE) AND  (x3 = FALSE) AND  ( TRUE ) AND  (x5 = TRUE)) OR ((x0 = TRUE) AND  ( TRUE ) AND  (x2 = FALSE) AND  (x3 = FALSE) AND  ( TRUE ) AND  (x5 = TRUE)) THEN 
        cstate98 := 1198; y0 := FALSE; y1 := FALSE; y2 := FALSE;  
    END_IF;
2696:
    IF ((x0 = FALSE) AND  (x1 = FALSE) AND  (x2 = FALSE) AND  ( TRUE ) AND  ( TRUE ) AND  (x5 = FALSE)) OR ((x0 = FALSE) AND  (x1 = TRUE) AND  (x2 = FALSE) AND  (x3 = FALSE) AND  ( TRUE ) AND  (x5 = FALSE)) OR ((x0 = TRUE) AND  ( TRUE ) AND  (x2 = FALSE) AND  (x3 = FALSE) AND  ( TRUE ) AND  (x5 = FALSE)) THEN 
        cstate98 := 3720; y0 := FALSE; y1 := TRUE; y2 := FALSE;  
    ELSIF ((x0 = FALSE) AND  (x1 = FALSE) AND  (x2 = FALSE) AND  (x3 = FALSE) AND  ( TRUE ) AND  (x5 = TRUE)) OR ((x0 = FALSE) AND  (x1 = FALSE) AND  (x2 = FALSE) AND  (x3 = TRUE) AND  (x4 = FALSE) AND  (x5 = TRUE)) THEN 
        cstate98 := 2219; y0 := FALSE; y1 := FALSE; y2 := FALSE;  
    ELSIF ((x0 = FALSE) AND  (x1 = FALSE) AND  (x2 = FALSE) AND  (x3 = TRUE) AND  (x4 = TRUE) AND  (x5 = TRUE)) THEN 
        cstate98 := 2186; y0 := FALSE; y1 := FALSE; y2 := FALSE;  
    ELSIF ((x0 = FALSE) AND  (x1 = FALSE) AND  (x2 = TRUE) AND  (x3 = FALSE) AND  ( TRUE ) AND  (x5 = FALSE)) THEN 
        cstate98 := 2696; y0 := FALSE; y1 := TRUE; y2 := FALSE;  
    ELSIF ((x0 = FALSE) AND  (x1 = FALSE) AND  (x2 = TRUE) AND  (x3 = FALSE) AND  ( TRUE ) AND  (x5 = TRUE)) THEN 
        cstate98 := 1706; y0 := FALSE; y1 := FALSE; y2 := FALSE;  
    ELSIF ((x0 = FALSE) AND  (x1 = FALSE) AND  (x2 = TRUE) AND  (x3 = TRUE) AND  ( TRUE ) AND  ( TRUE )) OR ((x0 = FALSE) AND  (x1 = TRUE) AND  (x2 = FALSE) AND  (x3 = TRUE) AND  ( TRUE ) AND  ( TRUE )) OR ((x0 = FALSE) AND  (x1 = TRUE) AND  (x2 = TRUE) AND  ( TRUE ) AND  ( TRUE ) AND  ( TRUE )) OR ((x0 = TRUE) AND  ( TRUE ) AND  (x2 = FALSE) AND  (x3 = TRUE) AND  ( TRUE ) AND  ( TRUE )) OR ((x0 = TRUE) AND  ( TRUE ) AND  (x2 = TRUE) AND  ( TRUE ) AND  ( TRUE ) AND  ( TRUE )) THEN 
        cstate98 := 617; y0 := FALSE; y1 := FALSE; y2 := FALSE;  
    ELSIF ((x0 = FALSE) AND  (x1 = TRUE) AND  (x2 = FALSE) AND  (x3 = FALSE) AND  ( TRUE ) AND  (x5 = TRUE)) OR ((x0 = TRUE) AND  ( TRUE ) AND  (x2 = FALSE) AND  (x3 = FALSE) AND  ( TRUE ) AND  (x5 = TRUE)) THEN 
        cstate98 := 1194; y0 := FALSE; y1 := FALSE; y2 := FALSE;  
    END_IF;
2223:
    IF ((x0 = FALSE) AND  (x1 = FALSE) AND  (x2 = FALSE) AND  (x3 = FALSE) AND  ( TRUE ) AND  ( TRUE )) OR ((x0 = FALSE) AND  (x1 = FALSE) AND  (x2 = FALSE) AND  (x3 = TRUE) AND  (x4 = FALSE) AND  ( TRUE )) THEN 
        cstate98 := 2223; y0 := FALSE; y1 := FALSE; y2 := FALSE;  
    ELSIF ((x0 = FALSE) AND  (x1 = FALSE) AND  (x2 = FALSE) AND  (x3 = TRUE) AND  (x4 = TRUE) AND  (x5 = FALSE)) THEN 
        cstate98 := 238; y0 := FALSE; y1 := FALSE; y2 := TRUE;  
    ELSIF ((x0 = FALSE) AND  (x1 = FALSE) AND  (x2 = FALSE) AND  (x3 = TRUE) AND  (x4 = TRUE) AND  (x5 = TRUE)) THEN 
        cstate98 := 2190; y0 := FALSE; y1 := FALSE; y2 := FALSE;  
    ELSIF ((x0 = FALSE) AND  (x1 = FALSE) AND  (x2 = TRUE) AND  (x3 = FALSE) AND  ( TRUE ) AND  (x5 = FALSE)) THEN 
        cstate98 := 2698; y0 := FALSE; y1 := TRUE; y2 := FALSE;  
    ELSIF ((x0 = FALSE) AND  (x1 = FALSE) AND  (x2 = TRUE) AND  (x3 = FALSE) AND  ( TRUE ) AND  (x5 = TRUE)) THEN 
        cstate98 := 1706; y0 := FALSE; y1 := FALSE; y2 := FALSE;  
    ELSIF ((x0 = FALSE) AND  (x1 = FALSE) AND  (x2 = TRUE) AND  (x3 = TRUE) AND  ( TRUE ) AND  ( TRUE )) OR ((x0 = FALSE) AND  (x1 = TRUE) AND  (x2 = FALSE) AND  (x3 = TRUE) AND  ( TRUE ) AND  ( TRUE )) OR ((x0 = FALSE) AND  (x1 = TRUE) AND  (x2 = TRUE) AND  ( TRUE ) AND  ( TRUE ) AND  ( TRUE )) OR ((x0 = TRUE) AND  ( TRUE ) AND  (x2 = FALSE) AND  (x3 = TRUE) AND  ( TRUE ) AND  ( TRUE )) OR ((x0 = TRUE) AND  ( TRUE ) AND  (x2 = TRUE) AND  ( TRUE ) AND  ( TRUE ) AND  ( TRUE )) THEN 
        cstate98 := 617; y0 := FALSE; y1 := FALSE; y2 := FALSE;  
    ELSIF ((x0 = FALSE) AND  (x1 = TRUE) AND  (x2 = FALSE) AND  (x3 = FALSE) AND  ( TRUE ) AND  (x5 = FALSE)) OR ((x0 = TRUE) AND  ( TRUE ) AND  (x2 = FALSE) AND  (x3 = FALSE) AND  ( TRUE ) AND  (x5 = FALSE)) THEN 
        cstate98 := 3214; y0 := TRUE; y1 := FALSE; y2 := FALSE;  
    ELSIF ((x0 = FALSE) AND  (x1 = TRUE) AND  (x2 = FALSE) AND  (x3 = FALSE) AND  ( TRUE ) AND  (x5 = TRUE)) OR ((x0 = TRUE) AND  ( TRUE ) AND  (x2 = FALSE) AND  (x3 = FALSE) AND  ( TRUE ) AND  (x5 = TRUE)) THEN 
        cstate98 := 1198; y0 := FALSE; y1 := FALSE; y2 := FALSE;  
    END_IF;
1706:
    IF ((x0 = FALSE) AND  (x1 = FALSE) AND  (x2 = FALSE) AND  (x3 = FALSE) AND  ( TRUE ) AND  (x5 = FALSE)) OR ((x0 = FALSE) AND  (x1 = FALSE) AND  (x2 = FALSE) AND  (x3 = TRUE) AND  (x4 = FALSE) AND  (x5 = FALSE)) THEN 
        cstate98 := 2218; y0 := FALSE; y1 := FALSE; y2 := FALSE;  
    ELSIF ((x0 = FALSE) AND  (x1 = FALSE) AND  (x2 = FALSE) AND  (x3 = FALSE) AND  ( TRUE ) AND  (x5 = TRUE)) OR ((x0 = FALSE) AND  (x1 = FALSE) AND  (x2 = FALSE) AND  (x3 = TRUE) AND  (x4 = FALSE) AND  (x5 = TRUE)) THEN 
        cstate98 := 2219; y0 := FALSE; y1 := FALSE; y2 := FALSE;  
    ELSIF ((x0 = FALSE) AND  (x1 = FALSE) AND  (x2 = FALSE) AND  (x3 = TRUE) AND  (x4 = TRUE) AND  (x5 = FALSE)) THEN 
        cstate98 := 234; y0 := FALSE; y1 := FALSE; y2 := TRUE;  
    ELSIF ((x0 = FALSE) AND  (x1 = FALSE) AND  (x2 = FALSE) AND  (x3 = TRUE) AND  (x4 = TRUE) AND  (x5 = TRUE)) THEN 
        cstate98 := 2186; y0 := FALSE; y1 := FALSE; y2 := FALSE;  
    ELSIF ((x0 = FALSE) AND  (x1 = FALSE) AND  (x2 = TRUE) AND  (x3 = FALSE) AND  ( TRUE ) AND  ( TRUE )) THEN 
        cstate98 := 1706; y0 := FALSE; y1 := FALSE; y2 := FALSE;  
    ELSIF ((x0 = FALSE) AND  (x1 = FALSE) AND  (x2 = TRUE) AND  (x3 = TRUE) AND  ( TRUE ) AND  ( TRUE )) OR ((x0 = FALSE) AND  (x1 = TRUE) AND  (x2 = FALSE) AND  (x3 = TRUE) AND  ( TRUE ) AND  ( TRUE )) OR ((x0 = FALSE) AND  (x1 = TRUE) AND  (x2 = TRUE) AND  ( TRUE ) AND  ( TRUE ) AND  ( TRUE )) OR ((x0 = TRUE) AND  ( TRUE ) AND  (x2 = FALSE) AND  (x3 = TRUE) AND  ( TRUE ) AND  ( TRUE )) OR ((x0 = TRUE) AND  ( TRUE ) AND  (x2 = TRUE) AND  ( TRUE ) AND  ( TRUE ) AND  ( TRUE )) THEN 
        cstate98 := 617; y0 := FALSE; y1 := FALSE; y2 := FALSE;  
    ELSIF ((x0 = FALSE) AND  (x1 = TRUE) AND  (x2 = FALSE) AND  (x3 = FALSE) AND  ( TRUE ) AND  (x5 = FALSE)) OR ((x0 = TRUE) AND  ( TRUE ) AND  (x2 = FALSE) AND  (x3 = FALSE) AND  ( TRUE ) AND  (x5 = FALSE)) THEN 
        cstate98 := 3210; y0 := TRUE; y1 := FALSE; y2 := FALSE;  
    ELSIF ((x0 = FALSE) AND  (x1 = TRUE) AND  (x2 = FALSE) AND  (x3 = FALSE) AND  ( TRUE ) AND  (x5 = TRUE)) OR ((x0 = TRUE) AND  ( TRUE ) AND  (x2 = FALSE) AND  (x3 = FALSE) AND  ( TRUE ) AND  (x5 = TRUE)) THEN 
        cstate98 := 1194; y0 := FALSE; y1 := FALSE; y2 := FALSE;  
    END_IF;
2226:
    IF ((x0 = FALSE) AND  (x1 = FALSE) AND  (x2 = FALSE) AND  (x3 = FALSE) AND  ( TRUE ) AND  (x5 = FALSE)) OR ((x0 = FALSE) AND  (x1 = FALSE) AND  (x2 = FALSE) AND  (x3 = TRUE) AND  (x4 = FALSE) AND  (x5 = FALSE)) THEN 
        cstate98 := 2226; y0 := FALSE; y1 := FALSE; y2 := FALSE;  
    ELSIF ((x0 = FALSE) AND  (x1 = FALSE) AND  (x2 = FALSE) AND  (x3 = FALSE) AND  ( TRUE ) AND  (x5 = TRUE)) OR ((x0 = FALSE) AND  (x1 = FALSE) AND  (x2 = FALSE) AND  (x3 = TRUE) AND  (x4 = FALSE) AND  (x5 = TRUE)) THEN 
        cstate98 := 2227; y0 := FALSE; y1 := FALSE; y2 := FALSE;  
    ELSIF ((x0 = FALSE) AND  (x1 = FALSE) AND  (x2 = FALSE) AND  (x3 = TRUE) AND  (x4 = TRUE) AND  (x5 = FALSE)) THEN 
        cstate98 := 234; y0 := FALSE; y1 := FALSE; y2 := TRUE;  
    ELSIF ((x0 = FALSE) AND  (x1 = FALSE) AND  (x2 = FALSE) AND  (x3 = TRUE) AND  (x4 = TRUE) AND  (x5 = TRUE)) THEN 
        cstate98 := 2186; y0 := FALSE; y1 := FALSE; y2 := FALSE;  
    ELSIF ((x0 = FALSE) AND  (x1 = FALSE) AND  (x2 = TRUE) AND  (x3 = FALSE) AND  ( TRUE ) AND  (x5 = FALSE)) THEN 
        cstate98 := 2706; y0 := FALSE; y1 := TRUE; y2 := FALSE;  
    ELSIF ((x0 = FALSE) AND  (x1 = FALSE) AND  (x2 = TRUE) AND  (x3 = FALSE) AND  ( TRUE ) AND  (x5 = TRUE)) THEN 
        cstate98 := 1714; y0 := FALSE; y1 := FALSE; y2 := FALSE;  
    ELSIF ((x0 = FALSE) AND  (x1 = FALSE) AND  (x2 = TRUE) AND  (x3 = TRUE) AND  ( TRUE ) AND  ( TRUE )) OR ((x0 = FALSE) AND  (x1 = TRUE) AND  (x2 = FALSE) AND  (x3 = TRUE) AND  ( TRUE ) AND  ( TRUE )) OR ((x0 = FALSE) AND  (x1 = TRUE) AND  (x2 = TRUE) AND  ( TRUE ) AND  ( TRUE ) AND  ( TRUE )) OR ((x0 = TRUE) AND  ( TRUE ) AND  (x2 = FALSE) AND  (x3 = TRUE) AND  ( TRUE ) AND  ( TRUE )) OR ((x0 = TRUE) AND  ( TRUE ) AND  (x2 = TRUE) AND  ( TRUE ) AND  ( TRUE ) AND  ( TRUE )) THEN 
        cstate98 := 617; y0 := FALSE; y1 := FALSE; y2 := FALSE;  
    ELSIF ((x0 = FALSE) AND  (x1 = TRUE) AND  (x2 = FALSE) AND  (x3 = FALSE) AND  ( TRUE ) AND  (x5 = FALSE)) OR ((x0 = TRUE) AND  ( TRUE ) AND  (x2 = FALSE) AND  (x3 = FALSE) AND  ( TRUE ) AND  (x5 = FALSE)) THEN 
        cstate98 := 3218; y0 := TRUE; y1 := FALSE; y2 := FALSE;  
    ELSIF ((x0 = FALSE) AND  (x1 = TRUE) AND  (x2 = FALSE) AND  (x3 = FALSE) AND  ( TRUE ) AND  (x5 = TRUE)) OR ((x0 = TRUE) AND  ( TRUE ) AND  (x2 = FALSE) AND  (x3 = FALSE) AND  ( TRUE ) AND  (x5 = TRUE)) THEN 
        cstate98 := 1202; y0 := FALSE; y1 := FALSE; y2 := FALSE;  
    END_IF;
2227:
    IF ((x0 = FALSE) AND  (x1 = FALSE) AND  (x2 = FALSE) AND  (x3 = FALSE) AND  ( TRUE ) AND  ( TRUE )) OR ((x0 = FALSE) AND  (x1 = FALSE) AND  (x2 = FALSE) AND  (x3 = TRUE) AND  (x4 = FALSE) AND  ( TRUE )) THEN 
        cstate98 := 2227; y0 := FALSE; y1 := FALSE; y2 := FALSE;  
    ELSIF ((x0 = FALSE) AND  (x1 = FALSE) AND  (x2 = FALSE) AND  (x3 = TRUE) AND  (x4 = TRUE) AND  (x5 = FALSE)) THEN 
        cstate98 := 234; y0 := FALSE; y1 := FALSE; y2 := TRUE;  
    ELSIF ((x0 = FALSE) AND  (x1 = FALSE) AND  (x2 = FALSE) AND  (x3 = TRUE) AND  (x4 = TRUE) AND  (x5 = TRUE)) THEN 
        cstate98 := 2186; y0 := FALSE; y1 := FALSE; y2 := FALSE;  
    ELSIF ((x0 = FALSE) AND  (x1 = FALSE) AND  (x2 = TRUE) AND  (x3 = FALSE) AND  ( TRUE ) AND  (x5 = FALSE)) THEN 
        cstate98 := 2706; y0 := FALSE; y1 := TRUE; y2 := FALSE;  
    ELSIF ((x0 = FALSE) AND  (x1 = FALSE) AND  (x2 = TRUE) AND  (x3 = FALSE) AND  ( TRUE ) AND  (x5 = TRUE)) THEN 
        cstate98 := 1714; y0 := FALSE; y1 := FALSE; y2 := FALSE;  
    ELSIF ((x0 = FALSE) AND  (x1 = FALSE) AND  (x2 = TRUE) AND  (x3 = TRUE) AND  ( TRUE ) AND  ( TRUE )) OR ((x0 = FALSE) AND  (x1 = TRUE) AND  (x2 = FALSE) AND  (x3 = TRUE) AND  ( TRUE ) AND  ( TRUE )) OR ((x0 = FALSE) AND  (x1 = TRUE) AND  (x2 = TRUE) AND  ( TRUE ) AND  ( TRUE ) AND  ( TRUE )) OR ((x0 = TRUE) AND  ( TRUE ) AND  (x2 = FALSE) AND  (x3 = TRUE) AND  ( TRUE ) AND  ( TRUE )) OR ((x0 = TRUE) AND  ( TRUE ) AND  (x2 = TRUE) AND  ( TRUE ) AND  ( TRUE ) AND  ( TRUE )) THEN 
        cstate98 := 617; y0 := FALSE; y1 := FALSE; y2 := FALSE;  
    ELSIF ((x0 = FALSE) AND  (x1 = TRUE) AND  (x2 = FALSE) AND  (x3 = FALSE) AND  ( TRUE ) AND  (x5 = FALSE)) OR ((x0 = TRUE) AND  ( TRUE ) AND  (x2 = FALSE) AND  (x3 = FALSE) AND  ( TRUE ) AND  (x5 = FALSE)) THEN 
        cstate98 := 3218; y0 := TRUE; y1 := FALSE; y2 := FALSE;  
    ELSIF ((x0 = FALSE) AND  (x1 = TRUE) AND  (x2 = FALSE) AND  (x3 = FALSE) AND  ( TRUE ) AND  (x5 = TRUE)) OR ((x0 = TRUE) AND  ( TRUE ) AND  (x2 = FALSE) AND  (x3 = FALSE) AND  ( TRUE ) AND  (x5 = TRUE)) THEN 
        cstate98 := 1202; y0 := FALSE; y1 := FALSE; y2 := FALSE;  
    END_IF;
4230:
    IF ((x0 = FALSE) AND  (x1 = FALSE) AND  (x2 = FALSE) AND  (x3 = FALSE) AND  ( TRUE ) AND  (x5 = FALSE)) OR ((x0 = FALSE) AND  (x1 = FALSE) AND  (x2 = FALSE) AND  (x3 = TRUE) AND  (x4 = FALSE) AND  (x5 = FALSE)) THEN 
        cstate98 := 4230; y0 := TRUE; y1 := FALSE; y2 := FALSE;  
    ELSIF ((x0 = FALSE) AND  (x1 = FALSE) AND  (x2 = FALSE) AND  (x3 = FALSE) AND  ( TRUE ) AND  (x5 = TRUE)) OR ((x0 = FALSE) AND  (x1 = FALSE) AND  (x2 = FALSE) AND  (x3 = TRUE) AND  (x4 = FALSE) AND  (x5 = TRUE)) THEN 
        cstate98 := 2215; y0 := FALSE; y1 := FALSE; y2 := FALSE;  
    ELSIF ((x0 = FALSE) AND  (x1 = FALSE) AND  (x2 = FALSE) AND  (x3 = TRUE) AND  (x4 = TRUE) AND  (x5 = FALSE)) THEN 
        cstate98 := 4238; y0 := TRUE; y1 := FALSE; y2 := FALSE;  
    ELSIF ((x0 = FALSE) AND  (x1 = FALSE) AND  (x2 = FALSE) AND  (x3 = TRUE) AND  (x4 = TRUE) AND  (x5 = TRUE)) THEN 
        cstate98 := 2190; y0 := FALSE; y1 := FALSE; y2 := FALSE;  
    ELSIF ((x0 = FALSE) AND  (x1 = FALSE) AND  (x2 = TRUE) AND  (x3 = FALSE) AND  ( TRUE ) AND  (x5 = FALSE)) THEN 
        cstate98 := 4242; y0 := TRUE; y1 := FALSE; y2 := FALSE;  
    ELSIF ((x0 = FALSE) AND  (x1 = FALSE) AND  (x2 = TRUE) AND  (x3 = FALSE) AND  ( TRUE ) AND  (x5 = TRUE)) THEN 
        cstate98 := 1714; y0 := FALSE; y1 := FALSE; y2 := FALSE;  
    ELSIF ((x0 = FALSE) AND  (x1 = FALSE) AND  (x2 = TRUE) AND  (x3 = TRUE) AND  ( TRUE ) AND  ( TRUE )) OR ((x0 = FALSE) AND  (x1 = TRUE) AND  (x2 = FALSE) AND  (x3 = TRUE) AND  ( TRUE ) AND  ( TRUE )) OR ((x0 = FALSE) AND  (x1 = TRUE) AND  (x2 = TRUE) AND  ( TRUE ) AND  ( TRUE ) AND  ( TRUE )) OR ((x0 = TRUE) AND  ( TRUE ) AND  (x2 = FALSE) AND  (x3 = TRUE) AND  ( TRUE ) AND  ( TRUE )) OR ((x0 = TRUE) AND  ( TRUE ) AND  (x2 = TRUE) AND  ( TRUE ) AND  ( TRUE ) AND  ( TRUE )) THEN 
        cstate98 := 617; y0 := FALSE; y1 := FALSE; y2 := FALSE;  
    ELSIF ((x0 = FALSE) AND  (x1 = TRUE) AND  (x2 = FALSE) AND  (x3 = FALSE) AND  ( TRUE ) AND  (x5 = FALSE)) OR ((x0 = TRUE) AND  ( TRUE ) AND  (x2 = FALSE) AND  (x3 = FALSE) AND  ( TRUE ) AND  (x5 = FALSE)) THEN 
        cstate98 := 3206; y0 := TRUE; y1 := FALSE; y2 := FALSE;  
    ELSIF ((x0 = FALSE) AND  (x1 = TRUE) AND  (x2 = FALSE) AND  (x3 = FALSE) AND  ( TRUE ) AND  (x5 = TRUE)) OR ((x0 = TRUE) AND  ( TRUE ) AND  (x2 = FALSE) AND  (x3 = FALSE) AND  ( TRUE ) AND  (x5 = TRUE)) THEN 
        cstate98 := 1190; y0 := FALSE; y1 := FALSE; y2 := FALSE;  
    END_IF;
2127:
    IF ((x0 = FALSE) AND  (x1 = FALSE) AND  (x2 = FALSE) AND  (x3 = FALSE) AND  ( TRUE ) AND  ( TRUE )) OR ((x0 = FALSE) AND  (x1 = FALSE) AND  (x2 = FALSE) AND  (x3 = TRUE) AND  (x4 = FALSE) AND  ( TRUE )) THEN 
        cstate98 := 2127; y0 := FALSE; y1 := FALSE; y2 := FALSE;  
    ELSIF ((x0 = FALSE) AND  (x1 = FALSE) AND  (x2 = FALSE) AND  (x3 = TRUE) AND  (x4 = TRUE) AND  (x5 = FALSE)) THEN 
        cstate98 := 206; y0 := FALSE; y1 := FALSE; y2 := TRUE;  
    ELSIF ((x0 = FALSE) AND  (x1 = FALSE) AND  (x2 = FALSE) AND  (x3 = TRUE) AND  (x4 = TRUE) AND  (x5 = TRUE)) THEN 
        cstate98 := 2094; y0 := FALSE; y1 := FALSE; y2 := FALSE;  
    ELSIF ((x0 = FALSE) AND  (x1 = FALSE) AND  (x2 = TRUE) AND  (x3 = FALSE) AND  ( TRUE ) AND  (x5 = FALSE)) THEN 
        cstate98 := 2602; y0 := FALSE; y1 := TRUE; y2 := FALSE;  
    ELSIF ((x0 = FALSE) AND  (x1 = FALSE) AND  (x2 = TRUE) AND  (x3 = FALSE) AND  ( TRUE ) AND  (x5 = TRUE)) THEN 
        cstate98 := 1610; y0 := FALSE; y1 := FALSE; y2 := FALSE;  
    ELSIF ((x0 = FALSE) AND  (x1 = FALSE) AND  (x2 = TRUE) AND  (x3 = TRUE) AND  ( TRUE ) AND  ( TRUE )) OR ((x0 = FALSE) AND  (x1 = TRUE) AND  (x2 = FALSE) AND  (x3 = TRUE) AND  ( TRUE ) AND  ( TRUE )) OR ((x0 = FALSE) AND  (x1 = TRUE) AND  (x2 = TRUE) AND  ( TRUE ) AND  ( TRUE ) AND  ( TRUE )) OR ((x0 = TRUE) AND  ( TRUE ) AND  (x2 = FALSE) AND  (x3 = TRUE) AND  ( TRUE ) AND  ( TRUE )) OR ((x0 = TRUE) AND  ( TRUE ) AND  (x2 = TRUE) AND  ( TRUE ) AND  ( TRUE ) AND  ( TRUE )) THEN 
        cstate98 := 617; y0 := FALSE; y1 := FALSE; y2 := FALSE;  
    ELSIF ((x0 = FALSE) AND  (x1 = TRUE) AND  (x2 = FALSE) AND  (x3 = FALSE) AND  ( TRUE ) AND  (x5 = FALSE)) OR ((x0 = TRUE) AND  ( TRUE ) AND  (x2 = FALSE) AND  (x3 = FALSE) AND  ( TRUE ) AND  (x5 = FALSE)) THEN 
        cstate98 := 3214; y0 := TRUE; y1 := FALSE; y2 := FALSE;  
    ELSIF ((x0 = FALSE) AND  (x1 = TRUE) AND  (x2 = FALSE) AND  (x3 = FALSE) AND  ( TRUE ) AND  (x5 = TRUE)) OR ((x0 = TRUE) AND  ( TRUE ) AND  (x2 = FALSE) AND  (x3 = FALSE) AND  ( TRUE ) AND  (x5 = TRUE)) THEN 
        cstate98 := 1198; y0 := FALSE; y1 := FALSE; y2 := FALSE;  
    END_IF;
2128:
    IF ((x0 = FALSE) AND  (x1 = FALSE) AND  (x2 = FALSE) AND  (x3 = FALSE) AND  ( TRUE ) AND  (x5 = FALSE)) OR ((x0 = FALSE) AND  (x1 = FALSE) AND  (x2 = FALSE) AND  (x3 = TRUE) AND  (x4 = FALSE) AND  (x5 = FALSE)) THEN 
        cstate98 := 2128; y0 := FALSE; y1 := FALSE; y2 := FALSE;  
    ELSIF ((x0 = FALSE) AND  (x1 = FALSE) AND  (x2 = FALSE) AND  (x3 = FALSE) AND  ( TRUE ) AND  (x5 = TRUE)) OR ((x0 = FALSE) AND  (x1 = FALSE) AND  (x2 = FALSE) AND  (x3 = TRUE) AND  (x4 = FALSE) AND  (x5 = TRUE)) THEN 
        cstate98 := 2131; y0 := FALSE; y1 := FALSE; y2 := FALSE;  
    ELSIF ((x0 = FALSE) AND  (x1 = FALSE) AND  (x2 = FALSE) AND  (x3 = TRUE) AND  (x4 = TRUE) AND  (x5 = FALSE)) THEN 
        cstate98 := 200; y0 := FALSE; y1 := FALSE; y2 := TRUE;  
    ELSIF ((x0 = FALSE) AND  (x1 = FALSE) AND  (x2 = FALSE) AND  (x3 = TRUE) AND  (x4 = TRUE) AND  (x5 = TRUE)) THEN 
        cstate98 := 2090; y0 := FALSE; y1 := FALSE; y2 := FALSE;  
    ELSIF ((x0 = FALSE) AND  (x1 = FALSE) AND  (x2 = TRUE) AND  (x3 = FALSE) AND  ( TRUE ) AND  (x5 = FALSE)) THEN 
        cstate98 := 2608; y0 := FALSE; y1 := TRUE; y2 := FALSE;  
    ELSIF ((x0 = FALSE) AND  (x1 = FALSE) AND  (x2 = TRUE) AND  (x3 = FALSE) AND  ( TRUE ) AND  (x5 = TRUE)) THEN 
        cstate98 := 1618; y0 := FALSE; y1 := FALSE; y2 := FALSE;  
    ELSIF ((x0 = FALSE) AND  (x1 = FALSE) AND  (x2 = TRUE) AND  (x3 = TRUE) AND  ( TRUE ) AND  ( TRUE )) OR ((x0 = FALSE) AND  (x1 = TRUE) AND  (x2 = FALSE) AND  (x3 = TRUE) AND  ( TRUE ) AND  ( TRUE )) OR ((x0 = FALSE) AND  (x1 = TRUE) AND  (x2 = TRUE) AND  ( TRUE ) AND  ( TRUE ) AND  ( TRUE )) OR ((x0 = TRUE) AND  ( TRUE ) AND  (x2 = FALSE) AND  (x3 = TRUE) AND  ( TRUE ) AND  ( TRUE )) OR ((x0 = TRUE) AND  ( TRUE ) AND  (x2 = TRUE) AND  ( TRUE ) AND  ( TRUE ) AND  ( TRUE )) THEN 
        cstate98 := 617; y0 := FALSE; y1 := FALSE; y2 := FALSE;  
    ELSIF ((x0 = FALSE) AND  (x1 = TRUE) AND  (x2 = FALSE) AND  (x3 = FALSE) AND  ( TRUE ) AND  (x5 = FALSE)) OR ((x0 = TRUE) AND  ( TRUE ) AND  (x2 = FALSE) AND  (x3 = FALSE) AND  ( TRUE ) AND  (x5 = FALSE)) THEN 
        cstate98 := 3216; y0 := TRUE; y1 := FALSE; y2 := FALSE;  
    ELSIF ((x0 = FALSE) AND  (x1 = TRUE) AND  (x2 = FALSE) AND  (x3 = FALSE) AND  ( TRUE ) AND  (x5 = TRUE)) OR ((x0 = TRUE) AND  ( TRUE ) AND  (x2 = FALSE) AND  (x3 = FALSE) AND  ( TRUE ) AND  (x5 = TRUE)) THEN 
        cstate98 := 1202; y0 := FALSE; y1 := FALSE; y2 := FALSE;  
    END_IF;
268:
    IF ((x0 = FALSE) AND  (x1 = FALSE) AND  (x2 = FALSE) AND  (x3 = FALSE) AND  ( TRUE ) AND  (x5 = FALSE)) OR ((x0 = FALSE) AND  (x1 = FALSE) AND  (x2 = FALSE) AND  (x3 = TRUE) AND  (x4 = FALSE) AND  (x5 = FALSE)) THEN 
        cstate98 := 268; y0 := FALSE; y1 := FALSE; y2 := TRUE;  
    ELSIF ((x0 = FALSE) AND  (x1 = FALSE) AND  (x2 = FALSE) AND  (x3 = FALSE) AND  ( TRUE ) AND  (x5 = TRUE)) OR ((x0 = FALSE) AND  (x1 = FALSE) AND  (x2 = FALSE) AND  (x3 = TRUE) AND  (x4 = FALSE) AND  (x5 = TRUE)) THEN 
        cstate98 := 2127; y0 := FALSE; y1 := FALSE; y2 := FALSE;  
    ELSIF ((x0 = FALSE) AND  (x1 = FALSE) AND  (x2 = FALSE) AND  (x3 = TRUE) AND  (x4 = TRUE) AND  (x5 = FALSE)) THEN 
        cstate98 := 204; y0 := FALSE; y1 := FALSE; y2 := TRUE;  
    ELSIF ((x0 = FALSE) AND  (x1 = FALSE) AND  (x2 = FALSE) AND  (x3 = TRUE) AND  (x4 = TRUE) AND  (x5 = TRUE)) THEN 
        cstate98 := 2094; y0 := FALSE; y1 := FALSE; y2 := FALSE;  
    ELSIF ((x0 = FALSE) AND  (x1 = FALSE) AND  (x2 = TRUE) AND  (x3 = FALSE) AND  ( TRUE ) AND  (x5 = FALSE)) THEN 
        cstate98 := 264; y0 := FALSE; y1 := FALSE; y2 := TRUE;  
    ELSIF ((x0 = FALSE) AND  (x1 = FALSE) AND  (x2 = TRUE) AND  (x3 = FALSE) AND  ( TRUE ) AND  (x5 = TRUE)) THEN 
        cstate98 := 1610; y0 := FALSE; y1 := FALSE; y2 := FALSE;  
    ELSIF ((x0 = FALSE) AND  (x1 = FALSE) AND  (x2 = TRUE) AND  (x3 = TRUE) AND  ( TRUE ) AND  ( TRUE )) OR ((x0 = FALSE) AND  (x1 = TRUE) AND  (x2 = FALSE) AND  (x3 = TRUE) AND  ( TRUE ) AND  ( TRUE )) OR ((x0 = FALSE) AND  (x1 = TRUE) AND  (x2 = TRUE) AND  ( TRUE ) AND  ( TRUE ) AND  ( TRUE )) OR ((x0 = TRUE) AND  ( TRUE ) AND  (x2 = FALSE) AND  (x3 = TRUE) AND  ( TRUE ) AND  ( TRUE )) OR ((x0 = TRUE) AND  ( TRUE ) AND  (x2 = TRUE) AND  ( TRUE ) AND  ( TRUE ) AND  ( TRUE )) THEN 
        cstate98 := 617; y0 := FALSE; y1 := FALSE; y2 := FALSE;  
    ELSIF ((x0 = FALSE) AND  (x1 = TRUE) AND  (x2 = FALSE) AND  (x3 = FALSE) AND  ( TRUE ) AND  (x5 = FALSE)) OR ((x0 = TRUE) AND  ( TRUE ) AND  (x2 = FALSE) AND  (x3 = FALSE) AND  ( TRUE ) AND  (x5 = FALSE)) THEN 
        cstate98 := 300; y0 := FALSE; y1 := FALSE; y2 := TRUE;  
    ELSIF ((x0 = FALSE) AND  (x1 = TRUE) AND  (x2 = FALSE) AND  (x3 = FALSE) AND  ( TRUE ) AND  (x5 = TRUE)) OR ((x0 = TRUE) AND  ( TRUE ) AND  (x2 = FALSE) AND  (x3 = FALSE) AND  ( TRUE ) AND  (x5 = TRUE)) THEN 
        cstate98 := 1198; y0 := FALSE; y1 := FALSE; y2 := FALSE;  
    END_IF;
4234:
    IF ((x0 = FALSE) AND  (x1 = FALSE) AND  (x2 = FALSE) AND  ( TRUE ) AND  ( TRUE ) AND  (x5 = FALSE)) OR ((x0 = FALSE) AND  (x1 = FALSE) AND  (x2 = TRUE) AND  (x3 = FALSE) AND  ( TRUE ) AND  (x5 = FALSE)) THEN 
        cstate98 := 4234; y0 := TRUE; y1 := FALSE; y2 := FALSE;  
    ELSIF ((x0 = FALSE) AND  (x1 = FALSE) AND  (x2 = FALSE) AND  (x3 = FALSE) AND  ( TRUE ) AND  (x5 = TRUE)) OR ((x0 = FALSE) AND  (x1 = FALSE) AND  (x2 = FALSE) AND  (x3 = TRUE) AND  (x4 = FALSE) AND  (x5 = TRUE)) THEN 
        cstate98 := 2219; y0 := FALSE; y1 := FALSE; y2 := FALSE;  
    ELSIF ((x0 = FALSE) AND  (x1 = FALSE) AND  (x2 = FALSE) AND  (x3 = TRUE) AND  (x4 = TRUE) AND  (x5 = TRUE)) THEN 
        cstate98 := 2186; y0 := FALSE; y1 := FALSE; y2 := FALSE;  
    ELSIF ((x0 = FALSE) AND  (x1 = FALSE) AND  (x2 = TRUE) AND  (x3 = FALSE) AND  ( TRUE ) AND  (x5 = TRUE)) THEN 
        cstate98 := 1706; y0 := FALSE; y1 := FALSE; y2 := FALSE;  
    ELSIF ((x0 = FALSE) AND  (x1 = FALSE) AND  (x2 = TRUE) AND  (x3 = TRUE) AND  ( TRUE ) AND  ( TRUE )) OR ((x0 = FALSE) AND  (x1 = TRUE) AND  (x2 = FALSE) AND  (x3 = TRUE) AND  ( TRUE ) AND  ( TRUE )) OR ((x0 = FALSE) AND  (x1 = TRUE) AND  (x2 = TRUE) AND  ( TRUE ) AND  ( TRUE ) AND  ( TRUE )) OR ((x0 = TRUE) AND  ( TRUE ) AND  (x2 = FALSE) AND  (x3 = TRUE) AND  ( TRUE ) AND  ( TRUE )) OR ((x0 = TRUE) AND  ( TRUE ) AND  (x2 = TRUE) AND  ( TRUE ) AND  ( TRUE ) AND  ( TRUE )) THEN 
        cstate98 := 617; y0 := FALSE; y1 := FALSE; y2 := FALSE;  
    ELSIF ((x0 = FALSE) AND  (x1 = TRUE) AND  (x2 = FALSE) AND  (x3 = FALSE) AND  ( TRUE ) AND  (x5 = FALSE)) OR ((x0 = TRUE) AND  ( TRUE ) AND  (x2 = FALSE) AND  (x3 = FALSE) AND  ( TRUE ) AND  (x5 = FALSE)) THEN 
        cstate98 := 3210; y0 := TRUE; y1 := FALSE; y2 := FALSE;  
    ELSIF ((x0 = FALSE) AND  (x1 = TRUE) AND  (x2 = FALSE) AND  (x3 = FALSE) AND  ( TRUE ) AND  (x5 = TRUE)) OR ((x0 = TRUE) AND  ( TRUE ) AND  (x2 = FALSE) AND  (x3 = FALSE) AND  ( TRUE ) AND  (x5 = TRUE)) THEN 
        cstate98 := 1194; y0 := FALSE; y1 := FALSE; y2 := FALSE;  
    END_IF;
2126:
    IF ((x0 = FALSE) AND  (x1 = FALSE) AND  (x2 = FALSE) AND  (x3 = FALSE) AND  ( TRUE ) AND  (x5 = FALSE)) OR ((x0 = FALSE) AND  (x1 = FALSE) AND  (x2 = FALSE) AND  (x3 = TRUE) AND  (x4 = FALSE) AND  (x5 = FALSE)) THEN 
        cstate98 := 2126; y0 := FALSE; y1 := FALSE; y2 := FALSE;  
    ELSIF ((x0 = FALSE) AND  (x1 = FALSE) AND  (x2 = FALSE) AND  (x3 = FALSE) AND  ( TRUE ) AND  (x5 = TRUE)) OR ((x0 = FALSE) AND  (x1 = FALSE) AND  (x2 = FALSE) AND  (x3 = TRUE) AND  (x4 = FALSE) AND  (x5 = TRUE)) THEN 
        cstate98 := 2127; y0 := FALSE; y1 := FALSE; y2 := FALSE;  
    ELSIF ((x0 = FALSE) AND  (x1 = FALSE) AND  (x2 = FALSE) AND  (x3 = TRUE) AND  (x4 = TRUE) AND  (x5 = FALSE)) THEN 
        cstate98 := 206; y0 := FALSE; y1 := FALSE; y2 := TRUE;  
    ELSIF ((x0 = FALSE) AND  (x1 = FALSE) AND  (x2 = FALSE) AND  (x3 = TRUE) AND  (x4 = TRUE) AND  (x5 = TRUE)) THEN 
        cstate98 := 2094; y0 := FALSE; y1 := FALSE; y2 := FALSE;  
    ELSIF ((x0 = FALSE) AND  (x1 = FALSE) AND  (x2 = TRUE) AND  (x3 = FALSE) AND  ( TRUE ) AND  (x5 = FALSE)) THEN 
        cstate98 := 2602; y0 := FALSE; y1 := TRUE; y2 := FALSE;  
    ELSIF ((x0 = FALSE) AND  (x1 = FALSE) AND  (x2 = TRUE) AND  (x3 = FALSE) AND  ( TRUE ) AND  (x5 = TRUE)) THEN 
        cstate98 := 1610; y0 := FALSE; y1 := FALSE; y2 := FALSE;  
    ELSIF ((x0 = FALSE) AND  (x1 = FALSE) AND  (x2 = TRUE) AND  (x3 = TRUE) AND  ( TRUE ) AND  ( TRUE )) OR ((x0 = FALSE) AND  (x1 = TRUE) AND  (x2 = FALSE) AND  (x3 = TRUE) AND  ( TRUE ) AND  ( TRUE )) OR ((x0 = FALSE) AND  (x1 = TRUE) AND  (x2 = TRUE) AND  ( TRUE ) AND  ( TRUE ) AND  ( TRUE )) OR ((x0 = TRUE) AND  ( TRUE ) AND  (x2 = FALSE) AND  (x3 = TRUE) AND  ( TRUE ) AND  ( TRUE )) OR ((x0 = TRUE) AND  ( TRUE ) AND  (x2 = TRUE) AND  ( TRUE ) AND  ( TRUE ) AND  ( TRUE )) THEN 
        cstate98 := 617; y0 := FALSE; y1 := FALSE; y2 := FALSE;  
    ELSIF ((x0 = FALSE) AND  (x1 = TRUE) AND  (x2 = FALSE) AND  (x3 = FALSE) AND  ( TRUE ) AND  (x5 = FALSE)) OR ((x0 = TRUE) AND  ( TRUE ) AND  (x2 = FALSE) AND  (x3 = FALSE) AND  ( TRUE ) AND  (x5 = FALSE)) THEN 
        cstate98 := 3214; y0 := TRUE; y1 := FALSE; y2 := FALSE;  
    ELSIF ((x0 = FALSE) AND  (x1 = TRUE) AND  (x2 = FALSE) AND  (x3 = FALSE) AND  ( TRUE ) AND  (x5 = TRUE)) OR ((x0 = TRUE) AND  ( TRUE ) AND  (x2 = FALSE) AND  (x3 = FALSE) AND  ( TRUE ) AND  (x5 = TRUE)) THEN 
        cstate98 := 1198; y0 := FALSE; y1 := FALSE; y2 := FALSE;  
    END_IF;
266:
    IF ((x0 = FALSE) AND  (x1 = FALSE) AND  (x2 = FALSE) AND  (x3 = FALSE) AND  ( TRUE ) AND  (x5 = FALSE)) OR ((x0 = FALSE) AND  (x1 = FALSE) AND  (x2 = FALSE) AND  (x3 = TRUE) AND  (x4 = FALSE) AND  (x5 = FALSE)) OR ((x0 = FALSE) AND  (x1 = FALSE) AND  (x2 = TRUE) AND  (x3 = FALSE) AND  ( TRUE ) AND  (x5 = FALSE)) THEN 
        cstate98 := 266; y0 := FALSE; y1 := FALSE; y2 := TRUE;  
    ELSIF ((x0 = FALSE) AND  (x1 = FALSE) AND  (x2 = FALSE) AND  (x3 = FALSE) AND  ( TRUE ) AND  (x5 = TRUE)) OR ((x0 = FALSE) AND  (x1 = FALSE) AND  (x2 = FALSE) AND  (x3 = TRUE) AND  (x4 = FALSE) AND  (x5 = TRUE)) THEN 
        cstate98 := 2123; y0 := FALSE; y1 := FALSE; y2 := FALSE;  
    ELSIF ((x0 = FALSE) AND  (x1 = FALSE) AND  (x2 = FALSE) AND  (x3 = TRUE) AND  (x4 = TRUE) AND  (x5 = FALSE)) THEN 
        cstate98 := 202; y0 := FALSE; y1 := FALSE; y2 := TRUE;  
    ELSIF ((x0 = FALSE) AND  (x1 = FALSE) AND  (x2 = FALSE) AND  (x3 = TRUE) AND  (x4 = TRUE) AND  (x5 = TRUE)) THEN 
        cstate98 := 2090; y0 := FALSE; y1 := FALSE; y2 := FALSE;  
    ELSIF ((x0 = FALSE) AND  (x1 = FALSE) AND  (x2 = TRUE) AND  (x3 = FALSE) AND  ( TRUE ) AND  (x5 = TRUE)) THEN 
        cstate98 := 1610; y0 := FALSE; y1 := FALSE; y2 := FALSE;  
    ELSIF ((x0 = FALSE) AND  (x1 = FALSE) AND  (x2 = TRUE) AND  (x3 = TRUE) AND  ( TRUE ) AND  ( TRUE )) OR ((x0 = FALSE) AND  (x1 = TRUE) AND  (x2 = FALSE) AND  (x3 = TRUE) AND  ( TRUE ) AND  ( TRUE )) OR ((x0 = FALSE) AND  (x1 = TRUE) AND  (x2 = TRUE) AND  ( TRUE ) AND  ( TRUE ) AND  ( TRUE )) OR ((x0 = TRUE) AND  ( TRUE ) AND  (x2 = FALSE) AND  (x3 = TRUE) AND  ( TRUE ) AND  ( TRUE )) OR ((x0 = TRUE) AND  ( TRUE ) AND  (x2 = TRUE) AND  ( TRUE ) AND  ( TRUE ) AND  ( TRUE )) THEN 
        cstate98 := 617; y0 := FALSE; y1 := FALSE; y2 := FALSE;  
    ELSIF ((x0 = FALSE) AND  (x1 = TRUE) AND  (x2 = FALSE) AND  (x3 = FALSE) AND  ( TRUE ) AND  (x5 = FALSE)) OR ((x0 = TRUE) AND  ( TRUE ) AND  (x2 = FALSE) AND  (x3 = FALSE) AND  ( TRUE ) AND  (x5 = FALSE)) THEN 
        cstate98 := 298; y0 := FALSE; y1 := FALSE; y2 := TRUE;  
    ELSIF ((x0 = FALSE) AND  (x1 = TRUE) AND  (x2 = FALSE) AND  (x3 = FALSE) AND  ( TRUE ) AND  (x5 = TRUE)) OR ((x0 = TRUE) AND  ( TRUE ) AND  (x2 = FALSE) AND  (x3 = FALSE) AND  ( TRUE ) AND  (x5 = TRUE)) THEN 
        cstate98 := 1194; y0 := FALSE; y1 := FALSE; y2 := FALSE;  
    END_IF;
4232:
    IF ((x0 = FALSE) AND  (x1 = FALSE) AND  (x2 = FALSE) AND  ( TRUE ) AND  ( TRUE ) AND  (x5 = FALSE)) OR ((x0 = FALSE) AND  (x1 = FALSE) AND  (x2 = TRUE) AND  (x3 = FALSE) AND  ( TRUE ) AND  (x5 = FALSE)) THEN 
        cstate98 := 4232; y0 := TRUE; y1 := FALSE; y2 := FALSE;  
    ELSIF ((x0 = FALSE) AND  (x1 = FALSE) AND  (x2 = FALSE) AND  (x3 = FALSE) AND  ( TRUE ) AND  (x5 = TRUE)) OR ((x0 = FALSE) AND  (x1 = FALSE) AND  (x2 = FALSE) AND  (x3 = TRUE) AND  (x4 = FALSE) AND  (x5 = TRUE)) THEN 
        cstate98 := 2219; y0 := FALSE; y1 := FALSE; y2 := FALSE;  
    ELSIF ((x0 = FALSE) AND  (x1 = FALSE) AND  (x2 = FALSE) AND  (x3 = TRUE) AND  (x4 = TRUE) AND  (x5 = TRUE)) THEN 
        cstate98 := 2186; y0 := FALSE; y1 := FALSE; y2 := FALSE;  
    ELSIF ((x0 = FALSE) AND  (x1 = FALSE) AND  (x2 = TRUE) AND  (x3 = FALSE) AND  ( TRUE ) AND  (x5 = TRUE)) THEN 
        cstate98 := 1706; y0 := FALSE; y1 := FALSE; y2 := FALSE;  
    ELSIF ((x0 = FALSE) AND  (x1 = FALSE) AND  (x2 = TRUE) AND  (x3 = TRUE) AND  ( TRUE ) AND  ( TRUE )) OR ((x0 = FALSE) AND  (x1 = TRUE) AND  (x2 = FALSE) AND  (x3 = TRUE) AND  ( TRUE ) AND  ( TRUE )) OR ((x0 = FALSE) AND  (x1 = TRUE) AND  (x2 = TRUE) AND  ( TRUE ) AND  ( TRUE ) AND  ( TRUE )) OR ((x0 = TRUE) AND  ( TRUE ) AND  (x2 = FALSE) AND  (x3 = TRUE) AND  ( TRUE ) AND  ( TRUE )) OR ((x0 = TRUE) AND  ( TRUE ) AND  (x2 = TRUE) AND  ( TRUE ) AND  ( TRUE ) AND  ( TRUE )) THEN 
        cstate98 := 617; y0 := FALSE; y1 := FALSE; y2 := FALSE;  
    ELSIF ((x0 = FALSE) AND  (x1 = TRUE) AND  (x2 = FALSE) AND  (x3 = FALSE) AND  ( TRUE ) AND  (x5 = FALSE)) OR ((x0 = TRUE) AND  ( TRUE ) AND  (x2 = FALSE) AND  (x3 = FALSE) AND  ( TRUE ) AND  (x5 = FALSE)) THEN 
        cstate98 := 3208; y0 := TRUE; y1 := FALSE; y2 := FALSE;  
    ELSIF ((x0 = FALSE) AND  (x1 = TRUE) AND  (x2 = FALSE) AND  (x3 = FALSE) AND  ( TRUE ) AND  (x5 = TRUE)) OR ((x0 = TRUE) AND  ( TRUE ) AND  (x2 = FALSE) AND  (x3 = FALSE) AND  ( TRUE ) AND  (x5 = TRUE)) THEN 
        cstate98 := 1194; y0 := FALSE; y1 := FALSE; y2 := FALSE;  
    END_IF;
2123:
    IF ((x0 = FALSE) AND  (x1 = FALSE) AND  (x2 = FALSE) AND  (x3 = FALSE) AND  ( TRUE ) AND  ( TRUE )) OR ((x0 = FALSE) AND  (x1 = FALSE) AND  (x2 = FALSE) AND  (x3 = TRUE) AND  (x4 = FALSE) AND  ( TRUE )) THEN 
        cstate98 := 2123; y0 := FALSE; y1 := FALSE; y2 := FALSE;  
    ELSIF ((x0 = FALSE) AND  (x1 = FALSE) AND  (x2 = FALSE) AND  (x3 = TRUE) AND  (x4 = TRUE) AND  (x5 = FALSE)) THEN 
        cstate98 := 202; y0 := FALSE; y1 := FALSE; y2 := TRUE;  
    ELSIF ((x0 = FALSE) AND  (x1 = FALSE) AND  (x2 = FALSE) AND  (x3 = TRUE) AND  (x4 = TRUE) AND  (x5 = TRUE)) THEN 
        cstate98 := 2090; y0 := FALSE; y1 := FALSE; y2 := FALSE;  
    ELSIF ((x0 = FALSE) AND  (x1 = FALSE) AND  (x2 = TRUE) AND  (x3 = FALSE) AND  ( TRUE ) AND  (x5 = FALSE)) THEN 
        cstate98 := 2602; y0 := FALSE; y1 := TRUE; y2 := FALSE;  
    ELSIF ((x0 = FALSE) AND  (x1 = FALSE) AND  (x2 = TRUE) AND  (x3 = FALSE) AND  ( TRUE ) AND  (x5 = TRUE)) THEN 
        cstate98 := 1610; y0 := FALSE; y1 := FALSE; y2 := FALSE;  
    ELSIF ((x0 = FALSE) AND  (x1 = FALSE) AND  (x2 = TRUE) AND  (x3 = TRUE) AND  ( TRUE ) AND  ( TRUE )) OR ((x0 = FALSE) AND  (x1 = TRUE) AND  (x2 = FALSE) AND  (x3 = TRUE) AND  ( TRUE ) AND  ( TRUE )) OR ((x0 = FALSE) AND  (x1 = TRUE) AND  (x2 = TRUE) AND  ( TRUE ) AND  ( TRUE ) AND  ( TRUE )) OR ((x0 = TRUE) AND  ( TRUE ) AND  (x2 = FALSE) AND  (x3 = TRUE) AND  ( TRUE ) AND  ( TRUE )) OR ((x0 = TRUE) AND  ( TRUE ) AND  (x2 = TRUE) AND  ( TRUE ) AND  ( TRUE ) AND  ( TRUE )) THEN 
        cstate98 := 617; y0 := FALSE; y1 := FALSE; y2 := FALSE;  
    ELSIF ((x0 = FALSE) AND  (x1 = TRUE) AND  (x2 = FALSE) AND  (x3 = FALSE) AND  ( TRUE ) AND  (x5 = FALSE)) OR ((x0 = TRUE) AND  ( TRUE ) AND  (x2 = FALSE) AND  (x3 = FALSE) AND  ( TRUE ) AND  (x5 = FALSE)) THEN 
        cstate98 := 3210; y0 := TRUE; y1 := FALSE; y2 := FALSE;  
    ELSIF ((x0 = FALSE) AND  (x1 = TRUE) AND  (x2 = FALSE) AND  (x3 = FALSE) AND  ( TRUE ) AND  (x5 = TRUE)) OR ((x0 = TRUE) AND  ( TRUE ) AND  (x2 = FALSE) AND  (x3 = FALSE) AND  ( TRUE ) AND  (x5 = TRUE)) THEN 
        cstate98 := 1194; y0 := FALSE; y1 := FALSE; y2 := FALSE;  
    END_IF;
2124:
    IF ((x0 = FALSE) AND  (x1 = FALSE) AND  (x2 = FALSE) AND  (x3 = FALSE) AND  ( TRUE ) AND  (x5 = FALSE)) OR ((x0 = FALSE) AND  (x1 = FALSE) AND  (x2 = FALSE) AND  (x3 = TRUE) AND  (x4 = FALSE) AND  (x5 = FALSE)) THEN 
        cstate98 := 2124; y0 := FALSE; y1 := FALSE; y2 := FALSE;  
    ELSIF ((x0 = FALSE) AND  (x1 = FALSE) AND  (x2 = FALSE) AND  (x3 = FALSE) AND  ( TRUE ) AND  (x5 = TRUE)) OR ((x0 = FALSE) AND  (x1 = FALSE) AND  (x2 = FALSE) AND  (x3 = TRUE) AND  (x4 = FALSE) AND  (x5 = TRUE)) THEN 
        cstate98 := 2127; y0 := FALSE; y1 := FALSE; y2 := FALSE;  
    ELSIF ((x0 = FALSE) AND  (x1 = FALSE) AND  (x2 = FALSE) AND  (x3 = TRUE) AND  (x4 = TRUE) AND  (x5 = FALSE)) THEN 
        cstate98 := 204; y0 := FALSE; y1 := FALSE; y2 := TRUE;  
    ELSIF ((x0 = FALSE) AND  (x1 = FALSE) AND  (x2 = FALSE) AND  (x3 = TRUE) AND  (x4 = TRUE) AND  (x5 = TRUE)) THEN 
        cstate98 := 2094; y0 := FALSE; y1 := FALSE; y2 := FALSE;  
    ELSIF ((x0 = FALSE) AND  (x1 = FALSE) AND  (x2 = TRUE) AND  (x3 = FALSE) AND  ( TRUE ) AND  (x5 = FALSE)) THEN 
        cstate98 := 2600; y0 := FALSE; y1 := TRUE; y2 := FALSE;  
    ELSIF ((x0 = FALSE) AND  (x1 = FALSE) AND  (x2 = TRUE) AND  (x3 = FALSE) AND  ( TRUE ) AND  (x5 = TRUE)) THEN 
        cstate98 := 1610; y0 := FALSE; y1 := FALSE; y2 := FALSE;  
    ELSIF ((x0 = FALSE) AND  (x1 = FALSE) AND  (x2 = TRUE) AND  (x3 = TRUE) AND  ( TRUE ) AND  ( TRUE )) OR ((x0 = FALSE) AND  (x1 = TRUE) AND  (x2 = FALSE) AND  (x3 = TRUE) AND  ( TRUE ) AND  ( TRUE )) OR ((x0 = FALSE) AND  (x1 = TRUE) AND  (x2 = TRUE) AND  ( TRUE ) AND  ( TRUE ) AND  ( TRUE )) OR ((x0 = TRUE) AND  ( TRUE ) AND  (x2 = FALSE) AND  (x3 = TRUE) AND  ( TRUE ) AND  ( TRUE )) OR ((x0 = TRUE) AND  ( TRUE ) AND  (x2 = TRUE) AND  ( TRUE ) AND  ( TRUE ) AND  ( TRUE )) THEN 
        cstate98 := 617; y0 := FALSE; y1 := FALSE; y2 := FALSE;  
    ELSIF ((x0 = FALSE) AND  (x1 = TRUE) AND  (x2 = FALSE) AND  (x3 = FALSE) AND  ( TRUE ) AND  (x5 = FALSE)) OR ((x0 = TRUE) AND  ( TRUE ) AND  (x2 = FALSE) AND  (x3 = FALSE) AND  ( TRUE ) AND  (x5 = FALSE)) THEN 
        cstate98 := 3212; y0 := TRUE; y1 := FALSE; y2 := FALSE;  
    ELSIF ((x0 = FALSE) AND  (x1 = TRUE) AND  (x2 = FALSE) AND  (x3 = FALSE) AND  ( TRUE ) AND  (x5 = TRUE)) OR ((x0 = TRUE) AND  ( TRUE ) AND  (x2 = FALSE) AND  (x3 = FALSE) AND  ( TRUE ) AND  (x5 = TRUE)) THEN 
        cstate98 := 1198; y0 := FALSE; y1 := FALSE; y2 := FALSE;  
    END_IF;
264:
    IF ((x0 = FALSE) AND  (x1 = FALSE) AND  (x2 = FALSE) AND  (x3 = FALSE) AND  ( TRUE ) AND  (x5 = FALSE)) OR ((x0 = FALSE) AND  (x1 = FALSE) AND  (x2 = FALSE) AND  (x3 = TRUE) AND  (x4 = FALSE) AND  (x5 = FALSE)) OR ((x0 = FALSE) AND  (x1 = FALSE) AND  (x2 = TRUE) AND  (x3 = FALSE) AND  ( TRUE ) AND  (x5 = FALSE)) THEN 
        cstate98 := 264; y0 := FALSE; y1 := FALSE; y2 := TRUE;  
    ELSIF ((x0 = FALSE) AND  (x1 = FALSE) AND  (x2 = FALSE) AND  (x3 = FALSE) AND  ( TRUE ) AND  (x5 = TRUE)) OR ((x0 = FALSE) AND  (x1 = FALSE) AND  (x2 = FALSE) AND  (x3 = TRUE) AND  (x4 = FALSE) AND  (x5 = TRUE)) THEN 
        cstate98 := 2123; y0 := FALSE; y1 := FALSE; y2 := FALSE;  
    ELSIF ((x0 = FALSE) AND  (x1 = FALSE) AND  (x2 = FALSE) AND  (x3 = TRUE) AND  (x4 = TRUE) AND  (x5 = FALSE)) THEN 
        cstate98 := 200; y0 := FALSE; y1 := FALSE; y2 := TRUE;  
    ELSIF ((x0 = FALSE) AND  (x1 = FALSE) AND  (x2 = FALSE) AND  (x3 = TRUE) AND  (x4 = TRUE) AND  (x5 = TRUE)) THEN 
        cstate98 := 2090; y0 := FALSE; y1 := FALSE; y2 := FALSE;  
    ELSIF ((x0 = FALSE) AND  (x1 = FALSE) AND  (x2 = TRUE) AND  (x3 = FALSE) AND  ( TRUE ) AND  (x5 = TRUE)) THEN 
        cstate98 := 1610; y0 := FALSE; y1 := FALSE; y2 := FALSE;  
    ELSIF ((x0 = FALSE) AND  (x1 = FALSE) AND  (x2 = TRUE) AND  (x3 = TRUE) AND  ( TRUE ) AND  ( TRUE )) OR ((x0 = FALSE) AND  (x1 = TRUE) AND  (x2 = FALSE) AND  (x3 = TRUE) AND  ( TRUE ) AND  ( TRUE )) OR ((x0 = FALSE) AND  (x1 = TRUE) AND  (x2 = TRUE) AND  ( TRUE ) AND  ( TRUE ) AND  ( TRUE )) OR ((x0 = TRUE) AND  ( TRUE ) AND  (x2 = FALSE) AND  (x3 = TRUE) AND  ( TRUE ) AND  ( TRUE )) OR ((x0 = TRUE) AND  ( TRUE ) AND  (x2 = TRUE) AND  ( TRUE ) AND  ( TRUE ) AND  ( TRUE )) THEN 
        cstate98 := 617; y0 := FALSE; y1 := FALSE; y2 := FALSE;  
    ELSIF ((x0 = FALSE) AND  (x1 = TRUE) AND  (x2 = FALSE) AND  (x3 = FALSE) AND  ( TRUE ) AND  (x5 = FALSE)) OR ((x0 = TRUE) AND  ( TRUE ) AND  (x2 = FALSE) AND  (x3 = FALSE) AND  ( TRUE ) AND  (x5 = FALSE)) THEN 
        cstate98 := 296; y0 := FALSE; y1 := FALSE; y2 := TRUE;  
    ELSIF ((x0 = FALSE) AND  (x1 = TRUE) AND  (x2 = FALSE) AND  (x3 = FALSE) AND  ( TRUE ) AND  (x5 = TRUE)) OR ((x0 = TRUE) AND  ( TRUE ) AND  (x2 = FALSE) AND  (x3 = FALSE) AND  ( TRUE ) AND  (x5 = TRUE)) THEN 
        cstate98 := 1194; y0 := FALSE; y1 := FALSE; y2 := FALSE;  
    END_IF;
3730:
    IF ((x0 = FALSE) AND  (x1 = FALSE) AND  (x2 = FALSE) AND  (x3 = FALSE) AND  ( TRUE ) AND  (x5 = FALSE)) OR ((x0 = FALSE) AND  (x1 = FALSE) AND  (x2 = FALSE) AND  (x3 = TRUE) AND  (x4 = FALSE) AND  (x5 = FALSE)) OR ((x0 = FALSE) AND  (x1 = TRUE) AND  (x2 = FALSE) AND  (x3 = FALSE) AND  ( TRUE ) AND  (x5 = FALSE)) OR ((x0 = TRUE) AND  ( TRUE ) AND  (x2 = FALSE) AND  (x3 = FALSE) AND  ( TRUE ) AND  (x5 = FALSE)) THEN 
        cstate98 := 3730; y0 := FALSE; y1 := TRUE; y2 := FALSE;  
    ELSIF ((x0 = FALSE) AND  (x1 = FALSE) AND  (x2 = FALSE) AND  (x3 = FALSE) AND  ( TRUE ) AND  (x5 = TRUE)) OR ((x0 = FALSE) AND  (x1 = FALSE) AND  (x2 = FALSE) AND  (x3 = TRUE) AND  (x4 = FALSE) AND  (x5 = TRUE)) THEN 
        cstate98 := 2227; y0 := FALSE; y1 := FALSE; y2 := FALSE;  
    ELSIF ((x0 = FALSE) AND  (x1 = FALSE) AND  (x2 = FALSE) AND  (x3 = TRUE) AND  (x4 = TRUE) AND  (x5 = FALSE)) THEN 
        cstate98 := 3722; y0 := FALSE; y1 := TRUE; y2 := FALSE;  
    ELSIF ((x0 = FALSE) AND  (x1 = FALSE) AND  (x2 = FALSE) AND  (x3 = TRUE) AND  (x4 = TRUE) AND  (x5 = TRUE)) THEN 
        cstate98 := 2186; y0 := FALSE; y1 := FALSE; y2 := FALSE;  
    ELSIF ((x0 = FALSE) AND  (x1 = FALSE) AND  (x2 = TRUE) AND  (x3 = FALSE) AND  ( TRUE ) AND  (x5 = FALSE)) THEN 
        cstate98 := 2706; y0 := FALSE; y1 := TRUE; y2 := FALSE;  
    ELSIF ((x0 = FALSE) AND  (x1 = FALSE) AND  (x2 = TRUE) AND  (x3 = FALSE) AND  ( TRUE ) AND  (x5 = TRUE)) THEN 
        cstate98 := 1714; y0 := FALSE; y1 := FALSE; y2 := FALSE;  
    ELSIF ((x0 = FALSE) AND  (x1 = FALSE) AND  (x2 = TRUE) AND  (x3 = TRUE) AND  ( TRUE ) AND  ( TRUE )) OR ((x0 = FALSE) AND  (x1 = TRUE) AND  (x2 = FALSE) AND  (x3 = TRUE) AND  ( TRUE ) AND  ( TRUE )) OR ((x0 = FALSE) AND  (x1 = TRUE) AND  (x2 = TRUE) AND  ( TRUE ) AND  ( TRUE ) AND  ( TRUE )) OR ((x0 = TRUE) AND  ( TRUE ) AND  (x2 = FALSE) AND  (x3 = TRUE) AND  ( TRUE ) AND  ( TRUE )) OR ((x0 = TRUE) AND  ( TRUE ) AND  (x2 = TRUE) AND  ( TRUE ) AND  ( TRUE ) AND  ( TRUE )) THEN 
        cstate98 := 617; y0 := FALSE; y1 := FALSE; y2 := FALSE;  
    ELSIF ((x0 = FALSE) AND  (x1 = TRUE) AND  (x2 = FALSE) AND  (x3 = FALSE) AND  ( TRUE ) AND  (x5 = TRUE)) OR ((x0 = TRUE) AND  ( TRUE ) AND  (x2 = FALSE) AND  (x3 = FALSE) AND  ( TRUE ) AND  (x5 = TRUE)) THEN 
        cstate98 := 1202; y0 := FALSE; y1 := FALSE; y2 := FALSE;  
    END_IF;
4236:
    IF ((x0 = FALSE) AND  (x1 = FALSE) AND  (x2 = FALSE) AND  ( TRUE ) AND  ( TRUE ) AND  (x5 = FALSE)) THEN 
        cstate98 := 4236; y0 := TRUE; y1 := FALSE; y2 := FALSE;  
    ELSIF ((x0 = FALSE) AND  (x1 = FALSE) AND  (x2 = FALSE) AND  (x3 = FALSE) AND  ( TRUE ) AND  (x5 = TRUE)) OR ((x0 = FALSE) AND  (x1 = FALSE) AND  (x2 = FALSE) AND  (x3 = TRUE) AND  (x4 = FALSE) AND  (x5 = TRUE)) THEN 
        cstate98 := 2223; y0 := FALSE; y1 := FALSE; y2 := FALSE;  
    ELSIF ((x0 = FALSE) AND  (x1 = FALSE) AND  (x2 = FALSE) AND  (x3 = TRUE) AND  (x4 = TRUE) AND  (x5 = TRUE)) THEN 
        cstate98 := 2190; y0 := FALSE; y1 := FALSE; y2 := FALSE;  
    ELSIF ((x0 = FALSE) AND  (x1 = FALSE) AND  (x2 = TRUE) AND  (x3 = FALSE) AND  ( TRUE ) AND  (x5 = FALSE)) THEN 
        cstate98 := 4232; y0 := TRUE; y1 := FALSE; y2 := FALSE;  
    ELSIF ((x0 = FALSE) AND  (x1 = FALSE) AND  (x2 = TRUE) AND  (x3 = FALSE) AND  ( TRUE ) AND  (x5 = TRUE)) THEN 
        cstate98 := 1706; y0 := FALSE; y1 := FALSE; y2 := FALSE;  
    ELSIF ((x0 = FALSE) AND  (x1 = FALSE) AND  (x2 = TRUE) AND  (x3 = TRUE) AND  ( TRUE ) AND  ( TRUE )) OR ((x0 = FALSE) AND  (x1 = TRUE) AND  (x2 = FALSE) AND  (x3 = TRUE) AND  ( TRUE ) AND  ( TRUE )) OR ((x0 = FALSE) AND  (x1 = TRUE) AND  (x2 = TRUE) AND  ( TRUE ) AND  ( TRUE ) AND  ( TRUE )) OR ((x0 = TRUE) AND  ( TRUE ) AND  (x2 = FALSE) AND  (x3 = TRUE) AND  ( TRUE ) AND  ( TRUE )) OR ((x0 = TRUE) AND  ( TRUE ) AND  (x2 = TRUE) AND  ( TRUE ) AND  ( TRUE ) AND  ( TRUE )) THEN 
        cstate98 := 617; y0 := FALSE; y1 := FALSE; y2 := FALSE;  
    ELSIF ((x0 = FALSE) AND  (x1 = TRUE) AND  (x2 = FALSE) AND  (x3 = FALSE) AND  ( TRUE ) AND  (x5 = FALSE)) OR ((x0 = TRUE) AND  ( TRUE ) AND  (x2 = FALSE) AND  (x3 = FALSE) AND  ( TRUE ) AND  (x5 = FALSE)) THEN 
        cstate98 := 3212; y0 := TRUE; y1 := FALSE; y2 := FALSE;  
    ELSIF ((x0 = FALSE) AND  (x1 = TRUE) AND  (x2 = FALSE) AND  (x3 = FALSE) AND  ( TRUE ) AND  (x5 = TRUE)) OR ((x0 = TRUE) AND  ( TRUE ) AND  (x2 = FALSE) AND  (x3 = FALSE) AND  ( TRUE ) AND  (x5 = TRUE)) THEN 
        cstate98 := 1198; y0 := FALSE; y1 := FALSE; y2 := FALSE;  
    END_IF;
4238:
    IF ((x0 = FALSE) AND  (x1 = FALSE) AND  (x2 = FALSE) AND  ( TRUE ) AND  ( TRUE ) AND  (x5 = FALSE)) THEN 
        cstate98 := 4238; y0 := TRUE; y1 := FALSE; y2 := FALSE;  
    ELSIF ((x0 = FALSE) AND  (x1 = FALSE) AND  (x2 = FALSE) AND  (x3 = FALSE) AND  ( TRUE ) AND  (x5 = TRUE)) OR ((x0 = FALSE) AND  (x1 = FALSE) AND  (x2 = FALSE) AND  (x3 = TRUE) AND  (x4 = FALSE) AND  (x5 = TRUE)) THEN 
        cstate98 := 2223; y0 := FALSE; y1 := FALSE; y2 := FALSE;  
    ELSIF ((x0 = FALSE) AND  (x1 = FALSE) AND  (x2 = FALSE) AND  (x3 = TRUE) AND  (x4 = TRUE) AND  (x5 = TRUE)) THEN 
        cstate98 := 2190; y0 := FALSE; y1 := FALSE; y2 := FALSE;  
    ELSIF ((x0 = FALSE) AND  (x1 = FALSE) AND  (x2 = TRUE) AND  (x3 = FALSE) AND  ( TRUE ) AND  (x5 = FALSE)) THEN 
        cstate98 := 4234; y0 := TRUE; y1 := FALSE; y2 := FALSE;  
    ELSIF ((x0 = FALSE) AND  (x1 = FALSE) AND  (x2 = TRUE) AND  (x3 = FALSE) AND  ( TRUE ) AND  (x5 = TRUE)) THEN 
        cstate98 := 1706; y0 := FALSE; y1 := FALSE; y2 := FALSE;  
    ELSIF ((x0 = FALSE) AND  (x1 = FALSE) AND  (x2 = TRUE) AND  (x3 = TRUE) AND  ( TRUE ) AND  ( TRUE )) OR ((x0 = FALSE) AND  (x1 = TRUE) AND  (x2 = FALSE) AND  (x3 = TRUE) AND  ( TRUE ) AND  ( TRUE )) OR ((x0 = FALSE) AND  (x1 = TRUE) AND  (x2 = TRUE) AND  ( TRUE ) AND  ( TRUE ) AND  ( TRUE )) OR ((x0 = TRUE) AND  ( TRUE ) AND  (x2 = FALSE) AND  (x3 = TRUE) AND  ( TRUE ) AND  ( TRUE )) OR ((x0 = TRUE) AND  ( TRUE ) AND  (x2 = TRUE) AND  ( TRUE ) AND  ( TRUE ) AND  ( TRUE )) THEN 
        cstate98 := 617; y0 := FALSE; y1 := FALSE; y2 := FALSE;  
    ELSIF ((x0 = FALSE) AND  (x1 = TRUE) AND  (x2 = FALSE) AND  (x3 = FALSE) AND  ( TRUE ) AND  (x5 = FALSE)) OR ((x0 = TRUE) AND  ( TRUE ) AND  (x2 = FALSE) AND  (x3 = FALSE) AND  ( TRUE ) AND  (x5 = FALSE)) THEN 
        cstate98 := 3214; y0 := TRUE; y1 := FALSE; y2 := FALSE;  
    ELSIF ((x0 = FALSE) AND  (x1 = TRUE) AND  (x2 = FALSE) AND  (x3 = FALSE) AND  ( TRUE ) AND  (x5 = TRUE)) OR ((x0 = TRUE) AND  ( TRUE ) AND  (x2 = FALSE) AND  (x3 = FALSE) AND  ( TRUE ) AND  (x5 = TRUE)) THEN 
        cstate98 := 1198; y0 := FALSE; y1 := FALSE; y2 := FALSE;  
    END_IF;
296:
    IF ((x0 = FALSE) AND  (x1 = FALSE) AND  (x2 = FALSE) AND  (x3 = FALSE) AND  ( TRUE ) AND  (x5 = FALSE)) OR ((x0 = FALSE) AND  (x1 = FALSE) AND  (x2 = FALSE) AND  (x3 = TRUE) AND  (x4 = FALSE) AND  (x5 = FALSE)) OR ((x0 = FALSE) AND  (x1 = FALSE) AND  (x2 = TRUE) AND  (x3 = FALSE) AND  ( TRUE ) AND  (x5 = FALSE)) OR ((x0 = FALSE) AND  (x1 = TRUE) AND  (x2 = FALSE) AND  (x3 = FALSE) AND  ( TRUE ) AND  (x5 = FALSE)) OR ((x0 = TRUE) AND  ( TRUE ) AND  (x2 = FALSE) AND  (x3 = FALSE) AND  ( TRUE ) AND  (x5 = FALSE)) THEN 
        cstate98 := 296; y0 := FALSE; y1 := FALSE; y2 := TRUE;  
    ELSIF ((x0 = FALSE) AND  (x1 = FALSE) AND  (x2 = FALSE) AND  (x3 = FALSE) AND  ( TRUE ) AND  (x5 = TRUE)) OR ((x0 = FALSE) AND  (x1 = FALSE) AND  (x2 = FALSE) AND  (x3 = TRUE) AND  (x4 = FALSE) AND  (x5 = TRUE)) THEN 
        cstate98 := 2219; y0 := FALSE; y1 := FALSE; y2 := FALSE;  
    ELSIF ((x0 = FALSE) AND  (x1 = FALSE) AND  (x2 = FALSE) AND  (x3 = TRUE) AND  (x4 = TRUE) AND  (x5 = FALSE)) THEN 
        cstate98 := 232; y0 := FALSE; y1 := FALSE; y2 := TRUE;  
    ELSIF ((x0 = FALSE) AND  (x1 = FALSE) AND  (x2 = FALSE) AND  (x3 = TRUE) AND  (x4 = TRUE) AND  (x5 = TRUE)) THEN 
        cstate98 := 2186; y0 := FALSE; y1 := FALSE; y2 := FALSE;  
    ELSIF ((x0 = FALSE) AND  (x1 = FALSE) AND  (x2 = TRUE) AND  (x3 = FALSE) AND  ( TRUE ) AND  (x5 = TRUE)) THEN 
        cstate98 := 1706; y0 := FALSE; y1 := FALSE; y2 := FALSE;  
    ELSIF ((x0 = FALSE) AND  (x1 = FALSE) AND  (x2 = TRUE) AND  (x3 = TRUE) AND  ( TRUE ) AND  ( TRUE )) OR ((x0 = FALSE) AND  (x1 = TRUE) AND  (x2 = FALSE) AND  (x3 = TRUE) AND  ( TRUE ) AND  ( TRUE )) OR ((x0 = FALSE) AND  (x1 = TRUE) AND  (x2 = TRUE) AND  ( TRUE ) AND  ( TRUE ) AND  ( TRUE )) OR ((x0 = TRUE) AND  ( TRUE ) AND  (x2 = FALSE) AND  (x3 = TRUE) AND  ( TRUE ) AND  ( TRUE )) OR ((x0 = TRUE) AND  ( TRUE ) AND  (x2 = TRUE) AND  ( TRUE ) AND  ( TRUE ) AND  ( TRUE )) THEN 
        cstate98 := 617; y0 := FALSE; y1 := FALSE; y2 := FALSE;  
    ELSIF ((x0 = FALSE) AND  (x1 = TRUE) AND  (x2 = FALSE) AND  (x3 = FALSE) AND  ( TRUE ) AND  (x5 = TRUE)) OR ((x0 = TRUE) AND  ( TRUE ) AND  (x2 = FALSE) AND  (x3 = FALSE) AND  ( TRUE ) AND  (x5 = TRUE)) THEN 
        cstate98 := 1194; y0 := FALSE; y1 := FALSE; y2 := FALSE;  
    END_IF;
298:
    IF ((x0 = FALSE) AND  (x1 = FALSE) AND  (x2 = FALSE) AND  (x3 = FALSE) AND  ( TRUE ) AND  (x5 = FALSE)) OR ((x0 = FALSE) AND  (x1 = FALSE) AND  (x2 = FALSE) AND  (x3 = TRUE) AND  (x4 = FALSE) AND  (x5 = FALSE)) OR ((x0 = FALSE) AND  (x1 = FALSE) AND  (x2 = TRUE) AND  (x3 = FALSE) AND  ( TRUE ) AND  (x5 = FALSE)) OR ((x0 = FALSE) AND  (x1 = TRUE) AND  (x2 = FALSE) AND  (x3 = FALSE) AND  ( TRUE ) AND  (x5 = FALSE)) OR ((x0 = TRUE) AND  ( TRUE ) AND  (x2 = FALSE) AND  (x3 = FALSE) AND  ( TRUE ) AND  (x5 = FALSE)) THEN 
        cstate98 := 298; y0 := FALSE; y1 := FALSE; y2 := TRUE;  
    ELSIF ((x0 = FALSE) AND  (x1 = FALSE) AND  (x2 = FALSE) AND  (x3 = FALSE) AND  ( TRUE ) AND  (x5 = TRUE)) OR ((x0 = FALSE) AND  (x1 = FALSE) AND  (x2 = FALSE) AND  (x3 = TRUE) AND  (x4 = FALSE) AND  (x5 = TRUE)) THEN 
        cstate98 := 2219; y0 := FALSE; y1 := FALSE; y2 := FALSE;  
    ELSIF ((x0 = FALSE) AND  (x1 = FALSE) AND  (x2 = FALSE) AND  (x3 = TRUE) AND  (x4 = TRUE) AND  (x5 = FALSE)) THEN 
        cstate98 := 234; y0 := FALSE; y1 := FALSE; y2 := TRUE;  
    ELSIF ((x0 = FALSE) AND  (x1 = FALSE) AND  (x2 = FALSE) AND  (x3 = TRUE) AND  (x4 = TRUE) AND  (x5 = TRUE)) THEN 
        cstate98 := 2186; y0 := FALSE; y1 := FALSE; y2 := FALSE;  
    ELSIF ((x0 = FALSE) AND  (x1 = FALSE) AND  (x2 = TRUE) AND  (x3 = FALSE) AND  ( TRUE ) AND  (x5 = TRUE)) THEN 
        cstate98 := 1706; y0 := FALSE; y1 := FALSE; y2 := FALSE;  
    ELSIF ((x0 = FALSE) AND  (x1 = FALSE) AND  (x2 = TRUE) AND  (x3 = TRUE) AND  ( TRUE ) AND  ( TRUE )) OR ((x0 = FALSE) AND  (x1 = TRUE) AND  (x2 = FALSE) AND  (x3 = TRUE) AND  ( TRUE ) AND  ( TRUE )) OR ((x0 = FALSE) AND  (x1 = TRUE) AND  (x2 = TRUE) AND  ( TRUE ) AND  ( TRUE ) AND  ( TRUE )) OR ((x0 = TRUE) AND  ( TRUE ) AND  (x2 = FALSE) AND  (x3 = TRUE) AND  ( TRUE ) AND  ( TRUE )) OR ((x0 = TRUE) AND  ( TRUE ) AND  (x2 = TRUE) AND  ( TRUE ) AND  ( TRUE ) AND  ( TRUE )) THEN 
        cstate98 := 617; y0 := FALSE; y1 := FALSE; y2 := FALSE;  
    ELSIF ((x0 = FALSE) AND  (x1 = TRUE) AND  (x2 = FALSE) AND  (x3 = FALSE) AND  ( TRUE ) AND  (x5 = TRUE)) OR ((x0 = TRUE) AND  ( TRUE ) AND  (x2 = FALSE) AND  (x3 = FALSE) AND  ( TRUE ) AND  (x5 = TRUE)) THEN 
        cstate98 := 1194; y0 := FALSE; y1 := FALSE; y2 := FALSE;  
    END_IF;
1202:
    IF ((x0 = FALSE) AND  (x1 = FALSE) AND  (x2 = FALSE) AND  (x3 = FALSE) AND  ( TRUE ) AND  (x5 = FALSE)) OR ((x0 = FALSE) AND  (x1 = FALSE) AND  (x2 = FALSE) AND  (x3 = TRUE) AND  (x4 = FALSE) AND  (x5 = FALSE)) THEN 
        cstate98 := 2226; y0 := FALSE; y1 := FALSE; y2 := FALSE;  
    ELSIF ((x0 = FALSE) AND  (x1 = FALSE) AND  (x2 = FALSE) AND  (x3 = FALSE) AND  ( TRUE ) AND  (x5 = TRUE)) OR ((x0 = FALSE) AND  (x1 = FALSE) AND  (x2 = FALSE) AND  (x3 = TRUE) AND  (x4 = FALSE) AND  (x5 = TRUE)) THEN 
        cstate98 := 2227; y0 := FALSE; y1 := FALSE; y2 := FALSE;  
    ELSIF ((x0 = FALSE) AND  (x1 = FALSE) AND  (x2 = FALSE) AND  (x3 = TRUE) AND  (x4 = TRUE) AND  (x5 = FALSE)) THEN 
        cstate98 := 234; y0 := FALSE; y1 := FALSE; y2 := TRUE;  
    ELSIF ((x0 = FALSE) AND  (x1 = FALSE) AND  (x2 = FALSE) AND  (x3 = TRUE) AND  (x4 = TRUE) AND  (x5 = TRUE)) THEN 
        cstate98 := 2186; y0 := FALSE; y1 := FALSE; y2 := FALSE;  
    ELSIF ((x0 = FALSE) AND  (x1 = FALSE) AND  (x2 = TRUE) AND  (x3 = FALSE) AND  ( TRUE ) AND  (x5 = FALSE)) THEN 
        cstate98 := 2706; y0 := FALSE; y1 := TRUE; y2 := FALSE;  
    ELSIF ((x0 = FALSE) AND  (x1 = FALSE) AND  (x2 = TRUE) AND  (x3 = FALSE) AND  ( TRUE ) AND  (x5 = TRUE)) THEN 
        cstate98 := 1714; y0 := FALSE; y1 := FALSE; y2 := FALSE;  
    ELSIF ((x0 = FALSE) AND  (x1 = FALSE) AND  (x2 = TRUE) AND  (x3 = TRUE) AND  ( TRUE ) AND  ( TRUE )) OR ((x0 = FALSE) AND  (x1 = TRUE) AND  (x2 = FALSE) AND  (x3 = TRUE) AND  ( TRUE ) AND  ( TRUE )) OR ((x0 = FALSE) AND  (x1 = TRUE) AND  (x2 = TRUE) AND  ( TRUE ) AND  ( TRUE ) AND  ( TRUE )) OR ((x0 = TRUE) AND  ( TRUE ) AND  (x2 = FALSE) AND  (x3 = TRUE) AND  ( TRUE ) AND  ( TRUE )) OR ((x0 = TRUE) AND  ( TRUE ) AND  (x2 = TRUE) AND  ( TRUE ) AND  ( TRUE ) AND  ( TRUE )) THEN 
        cstate98 := 617; y0 := FALSE; y1 := FALSE; y2 := FALSE;  
    ELSIF ((x0 = FALSE) AND  (x1 = TRUE) AND  (x2 = FALSE) AND  (x3 = FALSE) AND  ( TRUE ) AND  ( TRUE )) OR ((x0 = TRUE) AND  ( TRUE ) AND  (x2 = FALSE) AND  (x3 = FALSE) AND  ( TRUE ) AND  ( TRUE )) THEN 
        cstate98 := 1202; y0 := FALSE; y1 := FALSE; y2 := FALSE;  
    END_IF;
4240:
    IF ((x0 = FALSE) AND  (x1 = FALSE) AND  (x2 = FALSE) AND  (x3 = FALSE) AND  ( TRUE ) AND  (x5 = FALSE)) OR ((x0 = FALSE) AND  (x1 = FALSE) AND  (x2 = FALSE) AND  (x3 = TRUE) AND  (x4 = FALSE) AND  (x5 = FALSE)) OR ((x0 = FALSE) AND  (x1 = FALSE) AND  (x2 = TRUE) AND  (x3 = FALSE) AND  ( TRUE ) AND  (x5 = FALSE)) THEN 
        cstate98 := 4240; y0 := TRUE; y1 := FALSE; y2 := FALSE;  
    ELSIF ((x0 = FALSE) AND  (x1 = FALSE) AND  (x2 = FALSE) AND  (x3 = FALSE) AND  ( TRUE ) AND  (x5 = TRUE)) OR ((x0 = FALSE) AND  (x1 = FALSE) AND  (x2 = FALSE) AND  (x3 = TRUE) AND  (x4 = FALSE) AND  (x5 = TRUE)) THEN 
        cstate98 := 2227; y0 := FALSE; y1 := FALSE; y2 := FALSE;  
    ELSIF ((x0 = FALSE) AND  (x1 = FALSE) AND  (x2 = FALSE) AND  (x3 = TRUE) AND  (x4 = TRUE) AND  (x5 = FALSE)) THEN 
        cstate98 := 4232; y0 := TRUE; y1 := FALSE; y2 := FALSE;  
    ELSIF ((x0 = FALSE) AND  (x1 = FALSE) AND  (x2 = FALSE) AND  (x3 = TRUE) AND  (x4 = TRUE) AND  (x5 = TRUE)) THEN 
        cstate98 := 2186; y0 := FALSE; y1 := FALSE; y2 := FALSE;  
    ELSIF ((x0 = FALSE) AND  (x1 = FALSE) AND  (x2 = TRUE) AND  (x3 = FALSE) AND  ( TRUE ) AND  (x5 = TRUE)) THEN 
        cstate98 := 1714; y0 := FALSE; y1 := FALSE; y2 := FALSE;  
    ELSIF ((x0 = FALSE) AND  (x1 = FALSE) AND  (x2 = TRUE) AND  (x3 = TRUE) AND  ( TRUE ) AND  ( TRUE )) OR ((x0 = FALSE) AND  (x1 = TRUE) AND  (x2 = FALSE) AND  (x3 = TRUE) AND  ( TRUE ) AND  ( TRUE )) OR ((x0 = FALSE) AND  (x1 = TRUE) AND  (x2 = TRUE) AND  ( TRUE ) AND  ( TRUE ) AND  ( TRUE )) OR ((x0 = TRUE) AND  ( TRUE ) AND  (x2 = FALSE) AND  (x3 = TRUE) AND  ( TRUE ) AND  ( TRUE )) OR ((x0 = TRUE) AND  ( TRUE ) AND  (x2 = TRUE) AND  ( TRUE ) AND  ( TRUE ) AND  ( TRUE )) THEN 
        cstate98 := 617; y0 := FALSE; y1 := FALSE; y2 := FALSE;  
    ELSIF ((x0 = FALSE) AND  (x1 = TRUE) AND  (x2 = FALSE) AND  (x3 = FALSE) AND  ( TRUE ) AND  (x5 = FALSE)) OR ((x0 = TRUE) AND  ( TRUE ) AND  (x2 = FALSE) AND  (x3 = FALSE) AND  ( TRUE ) AND  (x5 = FALSE)) THEN 
        cstate98 := 3216; y0 := TRUE; y1 := FALSE; y2 := FALSE;  
    ELSIF ((x0 = FALSE) AND  (x1 = TRUE) AND  (x2 = FALSE) AND  (x3 = FALSE) AND  ( TRUE ) AND  (x5 = TRUE)) OR ((x0 = TRUE) AND  ( TRUE ) AND  (x2 = FALSE) AND  (x3 = FALSE) AND  ( TRUE ) AND  (x5 = TRUE)) THEN 
        cstate98 := 1202; y0 := FALSE; y1 := FALSE; y2 := FALSE;  
    END_IF;
2186:
    IF ((x0 = FALSE) AND  (x1 = FALSE) AND  (x2 = FALSE) AND  (x3 = FALSE) AND  ( TRUE ) AND  (x5 = FALSE)) OR ((x0 = FALSE) AND  (x1 = FALSE) AND  (x2 = FALSE) AND  (x3 = TRUE) AND  (x4 = FALSE) AND  (x5 = FALSE)) THEN 
        cstate98 := 2218; y0 := FALSE; y1 := FALSE; y2 := FALSE;  
    ELSIF ((x0 = FALSE) AND  (x1 = FALSE) AND  (x2 = FALSE) AND  (x3 = FALSE) AND  ( TRUE ) AND  (x5 = TRUE)) OR ((x0 = FALSE) AND  (x1 = FALSE) AND  (x2 = FALSE) AND  (x3 = TRUE) AND  (x4 = FALSE) AND  (x5 = TRUE)) THEN 
        cstate98 := 2219; y0 := FALSE; y1 := FALSE; y2 := FALSE;  
    ELSIF ((x0 = FALSE) AND  (x1 = FALSE) AND  (x2 = FALSE) AND  (x3 = TRUE) AND  (x4 = TRUE) AND  ( TRUE )) THEN 
        cstate98 := 2186; y0 := FALSE; y1 := FALSE; y2 := FALSE;  
    ELSIF ((x0 = FALSE) AND  (x1 = FALSE) AND  (x2 = TRUE) AND  (x3 = FALSE) AND  ( TRUE ) AND  (x5 = FALSE)) THEN 
        cstate98 := 2698; y0 := FALSE; y1 := TRUE; y2 := FALSE;  
    ELSIF ((x0 = FALSE) AND  (x1 = FALSE) AND  (x2 = TRUE) AND  (x3 = FALSE) AND  ( TRUE ) AND  (x5 = TRUE)) THEN 
        cstate98 := 1706; y0 := FALSE; y1 := FALSE; y2 := FALSE;  
    ELSIF ((x0 = FALSE) AND  (x1 = FALSE) AND  (x2 = TRUE) AND  (x3 = TRUE) AND  ( TRUE ) AND  ( TRUE )) OR ((x0 = FALSE) AND  (x1 = TRUE) AND  (x2 = FALSE) AND  (x3 = TRUE) AND  ( TRUE ) AND  ( TRUE )) OR ((x0 = FALSE) AND  (x1 = TRUE) AND  (x2 = TRUE) AND  ( TRUE ) AND  ( TRUE ) AND  ( TRUE )) OR ((x0 = TRUE) AND  ( TRUE ) AND  (x2 = FALSE) AND  (x3 = TRUE) AND  ( TRUE ) AND  ( TRUE )) OR ((x0 = TRUE) AND  ( TRUE ) AND  (x2 = TRUE) AND  ( TRUE ) AND  ( TRUE ) AND  ( TRUE )) THEN 
        cstate98 := 617; y0 := FALSE; y1 := FALSE; y2 := FALSE;  
    ELSIF ((x0 = FALSE) AND  (x1 = TRUE) AND  (x2 = FALSE) AND  (x3 = FALSE) AND  ( TRUE ) AND  (x5 = FALSE)) OR ((x0 = TRUE) AND  ( TRUE ) AND  (x2 = FALSE) AND  (x3 = FALSE) AND  ( TRUE ) AND  (x5 = FALSE)) THEN 
        cstate98 := 3210; y0 := TRUE; y1 := FALSE; y2 := FALSE;  
    ELSIF ((x0 = FALSE) AND  (x1 = TRUE) AND  (x2 = FALSE) AND  (x3 = FALSE) AND  ( TRUE ) AND  (x5 = TRUE)) OR ((x0 = TRUE) AND  ( TRUE ) AND  (x2 = FALSE) AND  (x3 = FALSE) AND  ( TRUE ) AND  (x5 = TRUE)) THEN 
        cstate98 := 1194; y0 := FALSE; y1 := FALSE; y2 := FALSE;  
    END_IF;
4242:
    IF ((x0 = FALSE) AND  (x1 = FALSE) AND  (x2 = FALSE) AND  (x3 = FALSE) AND  ( TRUE ) AND  (x5 = FALSE)) OR ((x0 = FALSE) AND  (x1 = FALSE) AND  (x2 = FALSE) AND  (x3 = TRUE) AND  (x4 = FALSE) AND  (x5 = FALSE)) OR ((x0 = FALSE) AND  (x1 = FALSE) AND  (x2 = TRUE) AND  (x3 = FALSE) AND  ( TRUE ) AND  (x5 = FALSE)) THEN 
        cstate98 := 4242; y0 := TRUE; y1 := FALSE; y2 := FALSE;  
    ELSIF ((x0 = FALSE) AND  (x1 = FALSE) AND  (x2 = FALSE) AND  (x3 = FALSE) AND  ( TRUE ) AND  (x5 = TRUE)) OR ((x0 = FALSE) AND  (x1 = FALSE) AND  (x2 = FALSE) AND  (x3 = TRUE) AND  (x4 = FALSE) AND  (x5 = TRUE)) THEN 
        cstate98 := 2227; y0 := FALSE; y1 := FALSE; y2 := FALSE;  
    ELSIF ((x0 = FALSE) AND  (x1 = FALSE) AND  (x2 = FALSE) AND  (x3 = TRUE) AND  (x4 = TRUE) AND  (x5 = FALSE)) THEN 
        cstate98 := 4234; y0 := TRUE; y1 := FALSE; y2 := FALSE;  
    ELSIF ((x0 = FALSE) AND  (x1 = FALSE) AND  (x2 = FALSE) AND  (x3 = TRUE) AND  (x4 = TRUE) AND  (x5 = TRUE)) THEN 
        cstate98 := 2186; y0 := FALSE; y1 := FALSE; y2 := FALSE;  
    ELSIF ((x0 = FALSE) AND  (x1 = FALSE) AND  (x2 = TRUE) AND  (x3 = FALSE) AND  ( TRUE ) AND  (x5 = TRUE)) THEN 
        cstate98 := 1714; y0 := FALSE; y1 := FALSE; y2 := FALSE;  
    ELSIF ((x0 = FALSE) AND  (x1 = FALSE) AND  (x2 = TRUE) AND  (x3 = TRUE) AND  ( TRUE ) AND  ( TRUE )) OR ((x0 = FALSE) AND  (x1 = TRUE) AND  (x2 = FALSE) AND  (x3 = TRUE) AND  ( TRUE ) AND  ( TRUE )) OR ((x0 = FALSE) AND  (x1 = TRUE) AND  (x2 = TRUE) AND  ( TRUE ) AND  ( TRUE ) AND  ( TRUE )) OR ((x0 = TRUE) AND  ( TRUE ) AND  (x2 = FALSE) AND  (x3 = TRUE) AND  ( TRUE ) AND  ( TRUE )) OR ((x0 = TRUE) AND  ( TRUE ) AND  (x2 = TRUE) AND  ( TRUE ) AND  ( TRUE ) AND  ( TRUE )) THEN 
        cstate98 := 617; y0 := FALSE; y1 := FALSE; y2 := FALSE;  
    ELSIF ((x0 = FALSE) AND  (x1 = TRUE) AND  (x2 = FALSE) AND  (x3 = FALSE) AND  ( TRUE ) AND  (x5 = FALSE)) OR ((x0 = TRUE) AND  ( TRUE ) AND  (x2 = FALSE) AND  (x3 = FALSE) AND  ( TRUE ) AND  (x5 = FALSE)) THEN 
        cstate98 := 3218; y0 := TRUE; y1 := FALSE; y2 := FALSE;  
    ELSIF ((x0 = FALSE) AND  (x1 = TRUE) AND  (x2 = FALSE) AND  (x3 = FALSE) AND  ( TRUE ) AND  (x5 = TRUE)) OR ((x0 = TRUE) AND  ( TRUE ) AND  (x2 = FALSE) AND  (x3 = FALSE) AND  ( TRUE ) AND  (x5 = TRUE)) THEN 
        cstate98 := 1202; y0 := FALSE; y1 := FALSE; y2 := FALSE;  
    END_IF;
617:
    IF ((x0 = FALSE) AND  (x1 = FALSE) AND  (x2 = FALSE) AND  ( TRUE ) AND  ( TRUE ) AND  ( TRUE )) OR ((x0 = FALSE) AND  (x1 = FALSE) AND  (x2 = TRUE) AND  (x3 = FALSE) AND  ( TRUE ) AND  ( TRUE )) OR ((x0 = FALSE) AND  (x1 = TRUE) AND  (x2 = FALSE) AND  (x3 = FALSE) AND  ( TRUE ) AND  ( TRUE )) OR ((x0 = TRUE) AND  ( TRUE ) AND  (x2 = FALSE) AND  (x3 = FALSE) AND  ( TRUE ) AND  ( TRUE )) THEN 
        cstate98 := 617; y0 := FALSE; y1 := FALSE; y2 := FALSE;  
    ELSIF ((x0 = FALSE) AND  (x1 = FALSE) AND  (x2 = TRUE) AND  (x3 = TRUE) AND  ( TRUE ) AND  ( TRUE )) OR ((x0 = FALSE) AND  (x1 = TRUE) AND  (x2 = FALSE) AND  (x3 = TRUE) AND  ( TRUE ) AND  ( TRUE )) OR ((x0 = FALSE) AND  (x1 = TRUE) AND  (x2 = TRUE) AND  ( TRUE ) AND  ( TRUE ) AND  ( TRUE )) OR ((x0 = TRUE) AND  ( TRUE ) AND  (x2 = FALSE) AND  (x3 = TRUE) AND  ( TRUE ) AND  ( TRUE )) OR ((x0 = TRUE) AND  ( TRUE ) AND  (x2 = TRUE) AND  ( TRUE ) AND  ( TRUE ) AND  ( TRUE )) THEN 
        cstate98 := 617; y0 := FALSE; y1 := FALSE; y2 := FALSE;  
    END_IF;
END_CASE;

END_FUNCTION_BLOCK
